       (*eDiagHistoryAbsolute*)
       1002:
         #Data.Parameter.Diag_History_Absolute.Power_Up_Counter.%B3:= #arrRecord[6];
         #Data.Parameter.Diag_History_Absolute.Power_Up_Counter.%B2:= #arrRecord[7];
         #Data.Parameter.Diag_History_Absolute.Power_Up_Counter.%B1:= #arrRecord[8];
         #Data.Parameter.Diag_History_Absolute.Power_Up_Counter.%B0:= #arrRecord[9];
         #Data.Parameter.Diag_History_Absolute.Operating_Time.%B3:= #arrRecord[10];
         #Data.Parameter.Diag_History_Absolute.Operating_Time.%B2:= #arrRecord[11];
         #Data.Parameter.Diag_History_Absolute.Operating_Time.%B1:= #arrRecord[12];
         #Data.Parameter.Diag_History_Absolute.Operating_Time.%B0:= #arrRecord[13];
         #Data.Parameter.Diag_History_Absolute.Maximum_Speed.%B3:= #arrRecord[14];
         #Data.Parameter.Diag_History_Absolute.Maximum_Speed.%B2:= #arrRecord[15];
         #Data.Parameter.Diag_History_Absolute.Maximum_Speed.%B1:= #arrRecord[16];
         #Data.Parameter.Diag_History_Absolute.Maximum_Speed.%B0:= #arrRecord[17];
         #Data.Parameter.Diag_History_Absolute.Counter_Rotation_fw.%B3:= #arrRecord[18];
         #Data.Parameter.Diag_History_Absolute.Counter_Rotation_fw.%B2:= #arrRecord[19];
         #Data.Parameter.Diag_History_Absolute.Counter_Rotation_fw.%B1:= #arrRecord[20];
         #Data.Parameter.Diag_History_Absolute.Counter_Rotation_fw.%B0:= #arrRecord[21];
         #Data.Parameter.Diag_History_Absolute.Counter_Rotation_bw.%B3:= #arrRecord[22];
         #Data.Parameter.Diag_History_Absolute.Counter_Rotation_bw.%B2:= #arrRecord[23];
         #Data.Parameter.Diag_History_Absolute.Counter_Rotation_bw.%B1:= #arrRecord[24];
         #Data.Parameter.Diag_History_Absolute.Counter_Rotation_bw.%B0:= #arrRecord[25];
         #Data.Parameter.Diag_History_Absolute.Counter_Rotation_alt.%B3:= #arrRecord[26];
         #Data.Parameter.Diag_History_Absolute.Counter_Rotation_alt.%B2:= #arrRecord[27];
         #Data.Parameter.Diag_History_Absolute.Counter_Rotation_alt.%B1:= #arrRecord[28];
         #Data.Parameter.Diag_History_Absolute.Counter_Rotation_alt.%B0:= #arrRecord[29];
         #Data.Parameter.Diag_History_Absolute.Counter_Motion.%B3:= #arrRecord[30];
         #Data.Parameter.Diag_History_Absolute.Counter_Motion.%B2:= #arrRecord[31];
         #Data.Parameter.Diag_History_Absolute.Counter_Motion.%B1:= #arrRecord[32];
         #Data.Parameter.Diag_History_Absolute.Counter_Motion.%B0:= #arrRecord[33];
         #Data.Parameter.Diag_History_Absolute.Reserved.%B3:= #arrRecord[34];
         #Data.Parameter.Diag_History_Absolute.Reserved.%B2:= #arrRecord[35];
         #Data.Parameter.Diag_History_Absolute.Reserved.%B1:= #arrRecord[36];
         #Data.Parameter.Diag_History_Absolute.Reserved.%B0:= #arrRecord[37];
         #Data.Parameter.Diag_History_Absolute.LED_Current_Maximum.%B3:= #arrRecord[38];
         #Data.Parameter.Diag_History_Absolute.LED_Current_Maximum.%B2:= #arrRecord[39];
         #Data.Parameter.Diag_History_Absolute.LED_Current_Maximum.%B1:= #arrRecord[40];
         #Data.Parameter.Diag_History_Absolute.LED_Current_Maximum.%B0:= #arrRecord[41];
         #Data.Parameter.Diag_History_Absolute.LED_Current_Minimum.%B3:= #arrRecord[42];
         #Data.Parameter.Diag_History_Absolute.LED_Current_Minimum.%B2:= #arrRecord[43];
         #Data.Parameter.Diag_History_Absolute.LED_Current_Minimum.%B1:= #arrRecord[44];
         #Data.Parameter.Diag_History_Absolute.LED_Current_Minimum.%B0:= #arrRecord[45];
         #Data.Parameter.Diag_History_Absolute.Voltage_Maximum.%B3:= #arrRecord[46];
         #Data.Parameter.Diag_History_Absolute.Voltage_Maximum.%B2:= #arrRecord[47];
         #Data.Parameter.Diag_History_Absolute.Voltage_Maximum.%B1:= #arrRecord[48];
         #Data.Parameter.Diag_History_Absolute.Voltage_Maximum.%B0:= #arrRecord[49];   
         #Data.Parameter.Diag_History_Absolute.Temperatur_Maximum.%B3:= #arrRecord[50];
         #Data.Parameter.Diag_History_Absolute.Temperatur_Maximum.%B2:= #arrRecord[51];
         #Data.Parameter.Diag_History_Absolute.Temperatur_Maximum.%B1:= #arrRecord[52];
         #Data.Parameter.Diag_History_Absolute.Temperatur_Maximum.%B0:= #arrRecord[53];
         #Data.Parameter.Diag_History_Absolute.Temperature_Minimum.%B3:= #arrRecord[54];
         #Data.Parameter.Diag_History_Absolute.Temperature_Minimum.%B2:= #arrRecord[55];
         #Data.Parameter.Diag_History_Absolute.Temperature_Minimum.%B1:= #arrRecord[56];
         #Data.Parameter.Diag_History_Absolute.Temperature_Minimum.%B0:= #arrRecord[57];

       (*eDiagHistoryRelative*)
       1003:
         #Data.Parameter.Diag_History_Relative.Power_Up_Counter.%B3:= #arrRecord[6];
         #Data.Parameter.Diag_History_Relative.Power_Up_Counter.%B2:= #arrRecord[7];
         #Data.Parameter.Diag_History_Relative.Power_Up_Counter.%B1:= #arrRecord[8];
         #Data.Parameter.Diag_History_Relative.Power_Up_Counter.%B0:= #arrRecord[9];
         #Data.Parameter.Diag_History_Relative.Operating_Time.%B3:= #arrRecord[10];
         #Data.Parameter.Diag_History_Relative.Operating_Time.%B2:= #arrRecord[11];
         #Data.Parameter.Diag_History_Relative.Operating_Time.%B1:= #arrRecord[12];
         #Data.Parameter.Diag_History_Relative.Operating_Time.%B0:= #arrRecord[13];
         #Data.Parameter.Diag_History_Relative.Maximum_Speed.%B3:= #arrRecord[14];
         #Data.Parameter.Diag_History_Relative.Maximum_Speed.%B2:= #arrRecord[15];
         #Data.Parameter.Diag_History_Relative.Maximum_Speed.%B1:= #arrRecord[16];
         #Data.Parameter.Diag_History_Relative.Maximum_Speed.%B0:= #arrRecord[17];
         #Data.Parameter.Diag_History_Relative.Counter_Rotation_fw.%B3:= #arrRecord[18];
         #Data.Parameter.Diag_History_Relative.Counter_Rotation_fw.%B2:= #arrRecord[19];
         #Data.Parameter.Diag_History_Relative.Counter_Rotation_fw.%B1:= #arrRecord[20];
         #Data.Parameter.Diag_History_Relative.Counter_Rotation_fw.%B0:= #arrRecord[21];
         #Data.Parameter.Diag_History_Relative.Counter_Rotation_bw.%B3:= #arrRecord[22];
         #Data.Parameter.Diag_History_Relative.Counter_Rotation_bw.%B2:= #arrRecord[23];
         #Data.Parameter.Diag_History_Relative.Counter_Rotation_bw.%B1:= #arrRecord[24];
         #Data.Parameter.Diag_History_Relative.Counter_Rotation_bw.%B0:= #arrRecord[25];
         #Data.Parameter.Diag_History_Relative.Counter_Rotation_alt.%B3:= #arrRecord[26];
         #Data.Parameter.Diag_History_Relative.Counter_Rotation_alt.%B2:= #arrRecord[27];
         #Data.Parameter.Diag_History_Relative.Counter_Rotation_alt.%B1:= #arrRecord[28];
         #Data.Parameter.Diag_History_Relative.Counter_Rotation_alt.%B0:= #arrRecord[29];
         #Data.Parameter.Diag_History_Relative.Counter_Motion.%B3:= #arrRecord[30];
         #Data.Parameter.Diag_History_Relative.Counter_Motion.%B2:= #arrRecord[31];
         #Data.Parameter.Diag_History_Relative.Counter_Motion.%B1:= #arrRecord[32];
         #Data.Parameter.Diag_History_Relative.Counter_Motion.%B0:= #arrRecord[33];
         #Data.Parameter.Diag_History_Relative.Reserved.%B3:= #arrRecord[34];
         #Data.Parameter.Diag_History_Relative.Reserved.%B2:= #arrRecord[35];
         #Data.Parameter.Diag_History_Relative.Reserved.%B1:= #arrRecord[36];
         #Data.Parameter.Diag_History_Relative.Reserved.%B0:= #arrRecord[37];
         #Data.Parameter.Diag_History_Relative.LED_Current_Maximum.%B3:= #arrRecord[38];
         #Data.Parameter.Diag_History_Relative.LED_Current_Maximum.%B2:= #arrRecord[39];
         #Data.Parameter.Diag_History_Relative.LED_Current_Maximum.%B1:= #arrRecord[40];
         #Data.Parameter.Diag_History_Relative.LED_Current_Maximum.%B0:= #arrRecord[41];
         #Data.Parameter.Diag_History_Relative.LED_Current_Minimum.%B3:= #arrRecord[42];
         #Data.Parameter.Diag_History_Relative.LED_Current_Minimum.%B2:= #arrRecord[43];
         #Data.Parameter.Diag_History_Relative.LED_Current_Minimum.%B1:= #arrRecord[44];
         #Data.Parameter.Diag_History_Relative.LED_Current_Minimum.%B0:= #arrRecord[45];
         #Data.Parameter.Diag_History_Relative.Voltage_Maximum.%B3:= #arrRecord[46];
         #Data.Parameter.Diag_History_Relative.Voltage_Maximum.%B2:= #arrRecord[47];
         #Data.Parameter.Diag_History_Relative.Voltage_Maximum.%B1:= #arrRecord[48];
         #Data.Parameter.Diag_History_Relative.Voltage_Maximum.%B0:= #arrRecord[49];   
         #Data.Parameter.Diag_History_Relative.Temperatur_Maximum.%B3:= #arrRecord[50];
         #Data.Parameter.Diag_History_Relative.Temperatur_Maximum.%B2:= #arrRecord[51];
         #Data.Parameter.Diag_History_Relative.Temperatur_Maximum.%B1:= #arrRecord[52];
         #Data.Parameter.Diag_History_Relative.Temperatur_Maximum.%B0:= #arrRecord[53];
         #Data.Parameter.Diag_History_Relative.Temperature_Minimum.%B3:= #arrRecord[54];
         #Data.Parameter.Diag_History_Relative.Temperature_Minimum.%B2:= #arrRecord[55];
         #Data.Parameter.Diag_History_Relative.Temperature_Minimum.%B1:= #arrRecord[56];
         #Data.Parameter.Diag_History_Relative.Temperature_Minimum.%B0:= #arrRecord[57];

       (*eDiagHistErrCounter*)
       1004:
         FOR #iIndex:= 0 TO 15 DO
           #Data.Parameter.Diag_Hist_Err_Counter[#iIndex].%B1:= #arrRecord[6 + 2 * #iIndex];
           #Data.Parameter.Diag_Hist_Err_Counter[#iIndex].%B0:= #arrRecord[7 + 2 * #iIndex];
         END_FOR;

       (*eSpeedCalculation*)
       1005:
         #Data.Parameter.Speed_Calculation.Control.%B1:= #arrRecord[6];
         #Data.Parameter.Speed_Calculation.Control.%B0:= #arrRecord[7];
         #Data.Parameter.Speed_Calculation.Velocity_Measuring_Unit.%B1:= #arrRecord[8];
         #Data.Parameter.Speed_Calculation.Velocity_Measuring_Unit.%B0:= #arrRecord[9];
         #Data.Parameter.Speed_Calculation.Update_Time_Tu.%B1:= #arrRecord[10];
         #Data.Parameter.Speed_Calculation.Update_Time_Tu.%B0:= #arrRecord[11];
         #Data.Parameter.Speed_Calculation.Update_Time_Ti.%B1:= #arrRecord[12];
         #Data.Parameter.Speed_Calculation.Update_Time_Ti.%B0:= #arrRecord[13];
         #Data.Parameter.Speed_Calculation.Upper_Limit.%B1:= #arrRecord[14];
         #Data.Parameter.Speed_Calculation.Upper_Limit.%B0:= #arrRecord[15];
         #Data.Parameter.Speed_Calculation.Lower_Limit.%B1:= #arrRecord[16];
         #Data.Parameter.Speed_Calculation.Lower_Limit.%B0:= #arrRecord[17];     

       (*eTemperatureLimits*)
       1006:
         #Data.Parameter.Temperature_Limits.Lower_Limit.%B1:= #arrRecord[6];
         #Data.Parameter.Temperature_Limits.Lower_Limit.%B0:= #arrRecord[7];
         #Data.Parameter.Temperature_Limits.Upper_Limit.%B1:= #arrRecord[8];
         #Data.Parameter.Temperature_Limits.Upper_Limit.%B0:= #arrRecord[9];   

       (*eVoltageLimits*)
       1007:
         #Data.Parameter.Voltage_Limits.Lower_Limit.%B1:= #arrRecord[6];
         #Data.Parameter.Voltage_Limits.Lower_Limit.%B0:= #arrRecord[7];
         #Data.Parameter.Voltage_Limits.Upper_Limit.%B1:= #arrRecord[8];
         #Data.Parameter.Voltage_Limits.Upper_Limit.%B0:= #arrRecord[9];   

       (*eScalingParameters*)
       1009: 
         #Data.Parameter.Scaling_Parameters.ES_Functionality.%B3:= #arrRecord[6];
         #Data.Parameter.Scaling_Parameters.ES_Functionality.%B2:= #arrRecord[7];
         #Data.Parameter.Scaling_Parameters.ES_Functionality.%B1:= #arrRecord[8];
         #Data.Parameter.Scaling_Parameters.ES_Functionality.%B0:= #arrRecord[9];
         #Data.Parameter.Scaling_Parameters.Input_CNR_N.%B3:= #arrRecord[10];
         #Data.Parameter.Scaling_Parameters.Input_CNR_N.%B2:= #arrRecord[11];
         #Data.Parameter.Scaling_Parameters.Input_CNR_N.%B1:= #arrRecord[12];
         #Data.Parameter.Scaling_Parameters.Input_CNR_N.%B0:= #arrRecord[13];
         #Data.Parameter.Scaling_Parameters.Input_CNR_D.%B3:= #arrRecord[14];
         #Data.Parameter.Scaling_Parameters.Input_CNR_D.%B2:= #arrRecord[15];
         #Data.Parameter.Scaling_Parameters.Input_CNR_D.%B1:= #arrRecord[16];
         #Data.Parameter.Scaling_Parameters.Input_CNR_D.%B0:= #arrRecord[17];
         #Data.Parameter.Scaling_Parameters.Input_CMR.%B3:= #arrRecord[18];
         #Data.Parameter.Scaling_Parameters.Input_CMR.%B2:= #arrRecord[19];
         #Data.Parameter.Scaling_Parameters.Input_CMR.%B1:= #arrRecord[20];
         #Data.Parameter.Scaling_Parameters.Input_CMR.%B0:= #arrRecord[21];
         #Data.Parameter.Scaling_Parameters.Range_Offset.%B3:= #arrRecord[22];
         #Data.Parameter.Scaling_Parameters.Range_Offset.%B2:= #arrRecord[23];
         #Data.Parameter.Scaling_Parameters.Range_Offset.%B1:= #arrRecord[24];
         #Data.Parameter.Scaling_Parameters.Range_Offset.%B0:= #arrRecord[25];
         #Data.Parameter.Scaling_Parameters.PMR_Shift.%B3:= #arrRecord[26];
         #Data.Parameter.Scaling_Parameters.PMR_Shift.%B2:= #arrRecord[27];
         #Data.Parameter.Scaling_Parameters.PMR_Shift.%B1:= #arrRecord[28];
         #Data.Parameter.Scaling_Parameters.PMR_Shift.%B0:= #arrRecord[29];
         #Data.Parameter.Scaling_Parameters.Output_CNR_N.%B3:= #arrRecord[30];
         #Data.Parameter.Scaling_Parameters.Output_CNR_N.%B2:= #arrRecord[31];
         #Data.Parameter.Scaling_Parameters.Output_CNR_N.%B1:= #arrRecord[32];
         #Data.Parameter.Scaling_Parameters.Output_CNR_N.%B0:= #arrRecord[33];
         #Data.Parameter.Scaling_Parameters.Output_CNR_D.%B3:= #arrRecord[34];
         #Data.Parameter.Scaling_Parameters.Output_CNR_D.%B2:= #arrRecord[35];
         #Data.Parameter.Scaling_Parameters.Output_CNR_D.%B1:= #arrRecord[36];
         #Data.Parameter.Scaling_Parameters.Output_CNR_D.%B0:= #arrRecord[37];
         #Data.Parameter.Scaling_Parameters.Output_CMR.%B3:= #arrRecord[38];
         #Data.Parameter.Scaling_Parameters.Output_CMR.%B2:= #arrRecord[39];
         #Data.Parameter.Scaling_Parameters.Output_CMR.%B1:= #arrRecord[40];
         #Data.Parameter.Scaling_Parameters.Output_CMR.%B0:= #arrRecord[41];
         #Data.Parameter.Scaling_Parameters.Out_CPR_Integer.%B3:= #arrRecord[42];
         #Data.Parameter.Scaling_Parameters.Out_CPR_Integer.%B2:= #arrRecord[43];
         #Data.Parameter.Scaling_Parameters.Out_CPR_Integer.%B1:= #arrRecord[44];
         #Data.Parameter.Scaling_Parameters.Out_CPR_Integer.%B0:= #arrRecord[45];
         #Data.Parameter.Scaling_Parameters.Out_CPR_Fract.%B3:= #arrRecord[46];
         #Data.Parameter.Scaling_Parameters.Out_CPR_Fract.%B2:= #arrRecord[47];
         #Data.Parameter.Scaling_Parameters.Out_CPR_Fract.%B1:= #arrRecord[48];
         #Data.Parameter.Scaling_Parameters.Out_CPR_Fract.%B0:= #arrRecord[49];

       (*eOperationTest1*)
       1010:
         #Data.Parameter.Operation_Test_1.%B1:= #arrRecord[6];
         #Data.Parameter.Operation_Test_1.%B0:= #arrRecord[7];

       (*eMACIDPort1*)
       1011:
         FOR #iIndex:= 0 TO 5 DO
           #Data.Parameter.MAC_ID_Port_1[#iIndex]:= #arrRecord[6 + #iIndex];
         END_FOR;

       (*eMACIDPort2*)
       1012:
         FOR #iIndex:= 0 TO 5 DO
           #Data.Parameter.MAC_ID_Port_2[#iIndex]:= #arrRecord[6 + #iIndex];
         END_FOR;

       (*eVersionFWFPGA*)
       1013:
         #Data.Parameter.Version_FW_FPGA.%B3:= #arrRecord[6];
         #Data.Parameter.Version_FW_FPGA.%B2:= #arrRecord[7];
         #Data.Parameter.Version_FW_FPGA.%B1:= #arrRecord[8];
         #Data.Parameter.Version_FW_FPGA.%B0:= #arrRecord[9];

       (*eTemperature*)
       1014:
         #Data.Parameter.Temperature.%B1:= #arrRecord[6];  
         #Data.Parameter.Temperature.%B0:= #arrRecord[7];  

       (*eStationName*)
       61000:
         Chars_TO_Strg(Chars:= #arrRecord, pChars:= 6, Cnt:= BYTE_TO_UINT(#arrRecord[5]), Strg=>#Data.Parameter.Station_Name);

       (*eStationIP*)
       61001:
         FOR #iIndex:= 0 TO 3 DO
           #Data.Parameter.Station_IP[#iIndex]:= #arrRecord[6 + #iIndex];
         END_FOR;

       (*eStationMACID*)
       61002:
         FOR #iIndex:= 0 TO 5 DO
           #Data.Parameter.Station_MAC_ID[#iIndex]:= #arrRecord[6 + #iIndex];
         END_FOR;

       (*eStationGateway*)
       61003:
         FOR #iIndex:= 0 TO 3 DO
           #Data.Parameter.Station_Gateway[#iIndex]:= #arrRecord[6 + #iIndex];
         END_FOR;

       (*eStationSubnet*)
       61004:
         FOR #iIndex:= 0 TO 3 DO
           #Data.Parameter.Station_Subnet[#iIndex]:= #arrRecord[6 + #iIndex];
         END_FOR;

       (*ePresetValue*)
       65000:
         #Data.Parameter.Preset_Value.%B3:= #arrRecord[6];
         #Data.Parameter.Preset_Value.%B2:= #arrRecord[7];
         #Data.Parameter.Preset_Value.%B1:= #arrRecord[8];
         #Data.Parameter.Preset_Value.%B0:= #arrRecord[9];

       (*eOperatingStatus*)
       65001:
         #Data.Parameter.Operating_Status.Header.%B3:= #arrRecord[6];
         #Data.Parameter.Operating_Status.Header.%B2:= #arrRecord[7];
         #Data.Parameter.Operating_Status.Header.%B1:= #arrRecord[8];
         #Data.Parameter.Operating_Status.Header.%B0:= #arrRecord[9];
         #Data.Parameter.Operating_Status.Operating_Status.%B3:= #arrRecord[10];
         #Data.Parameter.Operating_Status.Operating_Status.%B2:= #arrRecord[11];
         #Data.Parameter.Operating_Status.Operating_Status.%B1:= #arrRecord[12];
         #Data.Parameter.Operating_Status.Operating_Status.%B0:= #arrRecord[13];
         #Data.Parameter.Operating_Status.Faults.%B3:= #arrRecord[14];
         #Data.Parameter.Operating_Status.Faults.%B2:= #arrRecord[15];
         #Data.Parameter.Operating_Status.Faults.%B1:= #arrRecord[16];
         #Data.Parameter.Operating_Status.Faults.%B0:= #arrRecord[17];
         #Data.Parameter.Operating_Status.Supported_Faults.%B3:= #arrRecord[18];
         #Data.Parameter.Operating_Status.Supported_Faults.%B2:= #arrRecord[19];
         #Data.Parameter.Operating_Status.Supported_Faults.%B1:= #arrRecord[20];
         #Data.Parameter.Operating_Status.Supported_Faults.%B0:= #arrRecord[21];
         #Data.Parameter.Operating_Status.Warnings.%B3:= #arrRecord[22];
         #Data.Parameter.Operating_Status.Warnings.%B2:= #arrRecord[23];
         #Data.Parameter.Operating_Status.Warnings.%B1:= #arrRecord[24];
         #Data.Parameter.Operating_Status.Warnings.%B0:= #arrRecord[25];
         #Data.Parameter.Operating_Status.Supported_Warnings.%B3:= #arrRecord[26];
         #Data.Parameter.Operating_Status.Supported_Warnings.%B2:= #arrRecord[27];
         #Data.Parameter.Operating_Status.Supported_Warnings.%B1:= #arrRecord[28];
         #Data.Parameter.Operating_Status.Supported_Warnings.%B0:= #arrRecord[29];
         #Data.Parameter.Operating_Status.Encoder_Profile_Version.%B3:= #arrRecord[30];
         #Data.Parameter.Operating_Status.Encoder_Profile_Version.%B2:= #arrRecord[31];
         #Data.Parameter.Operating_Status.Encoder_Profile_Version.%B1:= #arrRecord[32];
         #Data.Parameter.Operating_Status.Encoder_Profile_Version.%B0:= #arrRecord[33];
         #Data.Parameter.Operating_Status.Operating_Time.%B3:= #arrRecord[34];
         #Data.Parameter.Operating_Status.Operating_Time.%B2:= #arrRecord[35];
         #Data.Parameter.Operating_Status.Operating_Time.%B1:= #arrRecord[36];
         #Data.Parameter.Operating_Status.Operating_Time.%B0:= #arrRecord[37];
         #Data.Parameter.Operating_Status.Offset_Value.%B3:= #arrRecord[38];
         #Data.Parameter.Operating_Status.Offset_Value.%B2:= #arrRecord[39];
         #Data.Parameter.Operating_Status.Offset_Value.%B1:= #arrRecord[40];
         #Data.Parameter.Operating_Status.Offset_Value.%B0:= #arrRecord[41];
         #Data.Parameter.Operating_Status.CPR.%B3:= #arrRecord[42];
         #Data.Parameter.Operating_Status.CPR.%B2:= #arrRecord[43];
         #Data.Parameter.Operating_Status.CPR.%B1:= #arrRecord[44];
         #Data.Parameter.Operating_Status.CPR.%B0:= #arrRecord[45];
         #Data.Parameter.Operating_Status.CMR.%B3:= #arrRecord[46];
         #Data.Parameter.Operating_Status.CMR.%B2:= #arrRecord[47];
         #Data.Parameter.Operating_Status.CMR.%B1:= #arrRecord[48];
         #Data.Parameter.Operating_Status.CMR.%B0:= #arrRecord[49];
         #Data.Parameter.Operating_Status.Velocity_Measuring_Unit.%B3:= #arrRecord[50];
         #Data.Parameter.Operating_Status.Velocity_Measuring_Unit.%B2:= #arrRecord[51];
         #Data.Parameter.Operating_Status.Velocity_Measuring_Unit.%B1:= #arrRecord[52];
         #Data.Parameter.Operating_Status.Velocity_Measuring_Unit.%B0:= #arrRecord[53];
     ELSE
       #stTempErrorCode.nBlockError:= 16#0002; (*Error: Internal error*)
     END_CASE;
     #iStep:= 9; (*Action permormed / Next command*)
   END_IF;


   (*======================== ACTION PERFORMED / NEXT COMMAND (STEP 9) =========================*)
   IF #iStep = 9 THEN
     #iCommandIndex:= #iCommandIndex + 1;

     (*Job done*)
     IF (#iCommandIndex > 31) OR (#arrCommandQueue[#iCommandIndex].iPNU <= 0) THEN
       #Done:= true;
       #Busy:= false;
       #bBusyMem:= false;
       #Error:= false;
       #iStep:= 0;

     (*Next command*)
     ELSE
       #iStep:= 4; (*Check communication status*)
     END_IF;
   END_IF;
END_FUNCTION_BLOCK

FUNCTION "Conveyors_Transfer" : Void   // FC24, SCL
{ S7_Optimized_Access := 'TRUE' }
VERSION : 0.1
// stored: AutoNumber true, IsIECCheckEnabled false, SetENOAutomatically false, UDAEnableTagReadback false
   VAR_TEMP
      i : Int;
   END_VAR
BEGIN
   //ID OF THE VTD CONVEYOR
   IF "Control_DB".VTD_Control.Current_Level = 0 THEN
       "Settings_DB".ECnv_Settings.ID := 120001;
       "Settings_DB".ECnv_Settings.Cnv_Level := 0;
   ELSIF "Control_DB".VTD_Control.Current_Level = 1 THEN
       "Settings_DB".ECnv_Settings.ID := 120101;
       "Settings_DB".ECnv_Settings.Cnv_Level := 1;
   ELSIF "Control_DB".VTD_Control.Current_Level = 2 THEN
       "Settings_DB".ECnv_Settings.ID := 120201;
       "Settings_DB".ECnv_Settings.Cnv_Level := 2;
   ELSIF "Control_DB".VTD_Control.Current_Level = 3 THEN
       "Settings_DB".ECnv_Settings.ID := 120301;
       "Settings_DB".ECnv_Settings.Cnv_Level := 3;
   ELSE
       "Settings_DB".ECnv_Settings.ID := 129901;
       "Settings_DB".ECnv_Settings.Cnv_Level := 99;
   END_IF;

   REGION READY TO RECEIVE
       //EXTRACTOR CONVEYOR
       "Control_DB".ECnv_Control.Instruction.Inbound_Ready :=
       ("Settings_DB".ECnv_Settings.ID = 120001 OR
       "Settings_DB".ECnv_Settings.ID = 120101 OR
       "Settings_DB".ECnv_Settings.ID = 120201 OR
       "Settings_DB".ECnv_Settings.ID = 120301)
       AND NOT "Control_DB".ECnv_Control.Cnv_Occupied AND NOT "Control_DB".ECnv_Control.Instruction.Outbound_Ready AND
       ("Control_DB".ECnv_Control.Mode = 2 OR "Control_DB".ECnv_Control.Mode = 3);

       //BUFFER CONVEYORS
       FOR #i := 1 TO 3 DO
           "Control_DB".LCnv_Control[#i].Instruction.Inbound_Ready :=
           NOT "Control_DB".LCnv_Control[#i].Running AND
           NOT "Control_DB".LCnv_Control[#i].Cnv_Occupied AND NOT "Control_DB".LCnv_Control[#i].Instruction.Outbound_Ready AND
           ("Control_DB".LCnv_Control[#i].Mode = 2 OR "Control_DB".LCnv_Control[#i].Mode = 3);
       END_FOR;

       //POPUP CONVEYORS
       FOR #i := 1 TO 4 DO
           "Control_DB".PopUp_Cnv[#i].Instruction.Inbound_Ready :=
           NOT "Control_DB".PopUp_Cnv[#i].Running AND
           NOT "Control_DB".PopUp_Cnv[#i].Cnv_Occupied AND NOT "Control_DB".PopUp_Cnv[#i].Instruction.Outbound_Ready AND
           ("Control_DB".PopUp_Cnv[#i].Mode = 2 OR "Control_DB".PopUp_Cnv[#i].Mode = 3);
       END_FOR;

       //INBOUND CONVEYOR
       "Control_DB".Inbound_Cnv.Instruction.Inbound_Ready := NOT "Control_DB".Inbound_Cnv.Cnv_Occupied;

       //OUTBOUND CONVEYOR
       "Control_DB".Outbound_Cnv.Instruction.Inbound_Ready :=
       NOT "Control_DB".Outbound_Cnv.Running AND
       NOT "Control_DB".Outbound_Cnv.Cnv_Occupied AND NOT "Control_DB".Outbound_Cnv.Instruction.Outbound_Ready AND
       ("Control_DB".Outbound_Cnv.Mode = 2 OR "Control_DB".Outbound_Cnv.Mode = 3);

       //PICK CONVEYOR
       "Control_DB".Pick_Station.Instruction.Inbound_Ready :=
       NOT "Control_DB".Pick_Station.Running AND
       NOT "Control_DB".Pick_Station.Cnv_Occupied AND NOT "Control_DB".Pick_Station.Instruction.Outbound_Ready AND
       ("Control_DB".Pick_Station.Mode = 2 OR "Control_DB".Pick_Station.Mode = 3);
   END_REGION

   REGION READY TO SEND
       //EXTRACTOR CONVEYOR
       "Control_DB".ECnv_Control.Instruction.Outbound_Ready :=
       (("Settings_DB".ECnv_Settings.ID = 120001 AND "Control_DB".ECnv_Control.Cnv_Occupied AND
       NOT "Control_DB".PopUp_Cnv[2].Cnv_Occupied AND ("Control_DB".PopUp_Cnv[2].Mode = 2 OR "Control_DB".PopUp_Cnv[2].Mode = 3)
       AND NOT "Control_DB".PopUp_Cnv[2].Error)
       OR
       ("Settings_DB".ECnv_Settings.ID = 120101 AND "Control_DB".ECnv_Control.Cnv_Occupied AND
       NOT "Control_DB".LCnv_Control[1].Cnv_Occupied AND ("Control_DB".LCnv_Control[1].Mode = 2 OR "Control_DB".LCnv_Control[1].Mode = 3)
       AND NOT "Control_DB".LCnv_Control[1].Error)
       OR
       ("Settings_DB".ECnv_Settings.ID = 120201 AND "Control_DB".ECnv_Control.Cnv_Occupied AND
       NOT "Control_DB".LCnv_Control[2].Cnv_Occupied AND ("Control_DB".LCnv_Control[2].Mode = 2 OR "Control_DB".LCnv_Control[2].Mode = 3)
       AND NOT "Control_DB".LCnv_Control[2].Error)
       OR
       ("Settings_DB".ECnv_Settings.ID = 120301 AND "Control_DB".ECnv_Control.Cnv_Occupied AND
       NOT "Control_DB".LCnv_Control[3].Cnv_Occupied AND ("Control_DB".LCnv_Control[3].Mode = 2 OR "Control_DB".LCnv_Control[3].Mode = 3)
       AND NOT "Control_DB".LCnv_Control[3].Error));

       //BUFFER CONVEYORS
       FOR #i := 1 TO 3 DO
           "Control_DB".LCnv_Control[#i].Instruction.Outbound_Ready :=
           "Control_DB".ECnv_Control.Instruction.Inbound_Ready AND
           "Control_DB".VTD_Control.Current_Level = #i AND
           NOT "Control_DB".LCnv_Control[#i].Instruction.Transfer_in_Progress AND
           "Control_DB".LCnv_Control[#i].Cnv_Occupied AND
           ("Control_DB".LCnv_Control[#i].Mode = 2 OR "Control_DB".LCnv_Control[#i].Mode = 3);
       END_FOR;

       //INBOUND CONVEYOR
       "Control_DB".Inbound_Cnv.Instruction.Outbound_Ready := "Control_DB".Inbound_Cnv.Cnv_Occupied;

       //POPUP CONVEYORS
       FOR #i := 1 TO 4 DO
           "Control_DB".PopUp_Cnv[#i].Instruction.Outbound_Ready :=
           ((#i = 1 AND "Control_DB".PopUp_Cnv[2].Instruction.Inbound_Ready AND "Control_DB".PopUp_Cnv[1].Inputs."Lift Up") OR
           (#i = 2 AND "Control_DB".PopUp_Cnv[2].Inputs."Lift Down" AND ("Control_DB".PopUp_Cnv[3].Instruction.Inbound_Ready OR "Control_DB".ECnv_Control.Instruction.Inbound_Ready)) OR
           (#i = 3 AND "Control_DB".PopUp_Cnv[4].Instruction.Inbound_Ready AND "Control_DB".PopUp_Cnv[3].Inputs."Lift Up") OR
           (#i = 4 AND ("Control_DB".Outbound_Cnv.Instruction.Inbound_Ready OR "Control_DB".PopUp_Cnv[1].Instruction.Inbound_Ready) AND ("Control_DB".PopUp_Cnv[4].Inputs."Lift Up" OR "Control_DB".PopUp_Cnv[4].Inputs."Lift Down"))) AND
           (*("Control_DB".VTD_Control.Current_Level = 0 AND #i = 2) AND*)
           NOT "Control_DB".PopUp_Cnv[#i].Instruction.Transfer_in_Progress AND
           "Control_DB".PopUp_Cnv[#i].Cnv_Occupied = TRUE AND
           ("Control_DB".PopUp_Cnv[#i].Mode = 2 OR "Control_DB".PopUp_Cnv[#i].Mode = 3);
       END_FOR;

       //PICK CONVEYOR
       "Control_DB".Pick_Station.Instruction.Outbound_Ready := "Control_DB".Pick_Station.Cnv_Occupied;
   END_REGION

   REGION TRANSFER IN PROGRESS FOR VTD
       "Cnv_TIP_For_VTD" :=
       ("Settings_DB".ECnv_Settings.ID = 120001 AND
       "Control_DB".PopUp_Cnv[2].Instruction.Transfer_in_Progress)
       OR
       ("Settings_DB".ECnv_Settings.ID = 120101 AND
       "Control_DB".LCnv_Control[1].Instruction.Transfer_in_Progress)
       OR
       ("Settings_DB".ECnv_Settings.ID = 120201 AND
       "Control_DB".LCnv_Control[2].Instruction.Transfer_in_Progress)
       OR
       ("Settings_DB".ECnv_Settings.ID = 120301 AND
       "Control_DB".LCnv_Control[3].Instruction.Transfer_in_Progress);
   END_REGION
END_FUNCTION

FUNCTION_BLOCK "Light_Bars"   // FB6, SCL
{ S7_Optimized_Access := 'TRUE' }
VERSION : 0.1
// stored: AutoNumber true, IsIECCheckEnabled false, IsRetainMemResEnabled false, MemoryReserve 100, SetENOAutomatically false, UDAEnableTagReadback false
   VAR_INPUT
      VTD_Mode : UInt;
      VTD_Speed : Int;
      Fault : Bool;
   END_VAR
   VAR_OUTPUT
      Animation_B1 : Byte;
      Color_B1 : Byte;
      Animation_B2 : Byte;
      Color_B2 : Byte;
      Speed_B1 : Byte;
      Speed_B2 : Byte;
   END_VAR
BEGIN
   //Commands for Light Bar

   IF #VTD_Mode = 0 AND NOT #Fault THEN // (0)Disabled = No light  
       #Animation_B1:= #Animation_B2:= 0;

   ELSIF #VTD_Mode = 1 AND #VTD_Speed = 0 AND  NOT #Fault AND NOT "SinaSpeed_VTD".EnableAxis THEN // (1)Manual= Yellow Stop
       #Animation_B1 := #Animation_B2 := 1;
       #Color_B1 := #Color_B2 := 4;

   ELSIF #VTD_Mode = 1 AND #VTD_Speed > 0 AND #VTD_Speed <= 33 AND  NOT #Fault AND "SinaSpeed_VTD".EnableAxis THEN // (1)Manual= Yellow until 33%
       #Animation_B1 := #Animation_B2 := 2;
       #Speed_B1 := #Speed_B2 := 2;
       #Color_B1 := #Color_B2 := 4;

   ELSIF #VTD_Mode = 1 AND #VTD_Speed > 33 AND #VTD_Speed <= 100 AND  NOT #Fault THEN // (1)Manual= Yellow until 66%
       #Animation_B1 := #Animation_B2 := 2;
       #Speed_B1 := #Speed_B2 := 0;
       #Color_B1 := #Color_B2 := 4;

   // ELSIF #VTD_Mode = 1 AND #VTD_Speed > 66 AND #VTD_Speed <= 100 AND  NOT #Fault THEN // (1)Manual= Yellow until 100%
   //     #Animation_B1 := #Animation_B2 := 2;
   //     #Speed_B1 := #Speed_B2 := 1;
   //     #Color_B1 := #Color_B2 := 4;

   ELSIF #VTD_Mode = 2 AND #VTD_Speed = 0 AND  NOT #Fault AND NOT "SinaSpeed_VTD".EnableAxis THEN // (2)Semi-auto = Blue Stop
       #Animation_B1 := #Animation_B2 := 1;
       #Color_B1 := #Color_B2 := 9;
       #Speed_B1 := #Speed_B2 := 0;

   ELSIF #VTD_Mode = 2 AND #VTD_Speed > 0 AND #VTD_Speed <= 33 AND  NOT #Fault AND "SinaSpeed_VTD".EnableAxis THEN // (2)Semi-auto = Blue until 33%
       #Animation_B1 := #Animation_B2 := 2;
       #Speed_B1 := #Speed_B2 := 2;
       #Color_B1 := #Color_B2 := 9;

   ELSIF #VTD_Mode = 2 AND #VTD_Speed > 33 AND #VTD_Speed <= 100 AND  NOT #Fault THEN // (2)Semi-auto = Blue until 66%
       #Animation_B1 := #Animation_B2 := 2;
       #Speed_B1 := #Speed_B2 := 0;
       #Color_B1 := #Color_B2 := 9;

   // ELSIF #VTD_Mode = 2 AND #VTD_Speed > 66 AND #VTD_Speed <= 100 AND  NOT #Fault THEN // (2)Semi-auto = Blue until 100%
   //     #Animation_B1 := #Animation_B2 := 2;
   //     #Speed_B1 := #Speed_B2 := 1;
   //     #Color_B1 := #Color_B2 := 9;

   ELSIF #VTD_Mode = 3 AND #VTD_Speed = 0 AND  NOT #Fault AND NOT "SinaSpeed_VTD".EnableAxis THEN // (3)Auto = Green Stop
       #Animation_B1 := #Animation_B2 := 1;
       #Color_B1 := #Color_B2 := 0;

   ELSIF #VTD_Mode = 3 AND #VTD_Speed > 0 AND #VTD_Speed <= 33 AND  NOT #Fault AND "SinaSpeed_VTD".EnableAxis THEN // (3)Auto = Green until 33%
       #Animation_B1 := #Animation_B2 := 2;
       #Speed_B1 := #Speed_B2 := 2;
       #Color_B1 := #Color_B2 := 0;

   ELSIF #VTD_Mode = 3 AND #VTD_Speed > 33 AND #VTD_Speed <= 100 AND  NOT #Fault THEN // (3)Auto = Green until 66%
       #Animation_B1 := #Animation_B2 := 2;
       #Speed_B1 := #Speed_B2 := 0;
       #Color_B1 := #Color_B2 := 0;

   // ELSIF #VTD_Mode = 3 AND #VTD_Speed > 66 AND #VTD_Speed <= 100 AND  NOT #Fault THEN // (3)Auto = Green until 100%
   //     #Animation_B1 := #Animation_B2 := 2;
   //     #Speed_B1 := #Speed_B2 := 1;
   //     #Color_B1 := #Color_B2 := 0;

   ELSIF #VTD_Mode = 4 AND #VTD_Speed = 0 AND  NOT #Fault THEN // (4)Tech = Orange Stop
       #Animation_B1 := #Animation_B2 := 1;
       #Color_B1 := #Color_B2 := 2;

   ELSIF #VTD_Mode = 4 AND #VTD_Speed > 0 AND #VTD_Speed <= 33 AND  NOT #Fault THEN // (4)Tech = Orange until 33%
       #Animation_B1 := #Animation_B2 := 2;
       #Speed_B1 := #Speed_B2 := 2;
       #Color_B1 := #Color_B2 := 2;

   ELSIF #VTD_Mode = 4 AND #VTD_Speed > 33 AND #VTD_Speed <= 66 AND  NOT #Fault THEN // (4)Tech = Orange until 66%
       #Animation_B1 := #Animation_B2 := 2;
       #Speed_B1 := #Speed_B2 := 0;
       #Color_B1 := #Color_B2 := 2;

   ELSIF #VTD_Mode = 4 AND #VTD_Speed > 66 AND #VTD_Speed <= 100 AND  NOT #Fault THEN // (4)Tech = Orange until 100%
       #Animation_B1 := #Animation_B2 := 2;
       #Speed_B1 := #Speed_B2 := 1;
       #Color_B1 := #Color_B2 := 2;

   ELSIF #VTD_Mode = 5 AND #VTD_Speed = 0 AND  NOT #Fault THEN // (5)Maintenance = White Stop
       #Animation_B1 := #Animation_B2 := 1;
       #Color_B1 := #Color_B2 := 19;

   ELSIF #VTD_Mode = 5 AND #VTD_Speed > 0 AND #VTD_Speed <= 33 AND  NOT #Fault THEN // (5)Maintenance = White until 33%
       #Animation_B1 := #Animation_B2 := 2;
       #Speed_B1 := #Speed_B2 := 2;
       #Color_B1 := #Color_B2 := 19;

   ELSIF #VTD_Mode = 5 AND #VTD_Speed > 33 AND #VTD_Speed <= 66 AND  NOT #Fault THEN // (5)Maintenance = White until 66%
       #Animation_B1 := #Animation_B2 := 2;
       #Speed_B1 := #Speed_B2 := 0;
       #Color_B1 := #Color_B2 := 19;

   ELSIF #VTD_Mode = 5 AND #VTD_Speed > 66 AND #VTD_Speed <= 100 AND  NOT #Fault THEN // (5)Maintenance = White until 100%
       #Animation_B1 := #Animation_B2 := 2;
       #Speed_B1 := #Speed_B2 := 1;
       #Color_B1 := #Color_B2 := 19;

   ELSIF #Fault THEN // Fault = Flash Red
       #Animation_B1:= #Animation_B2 := 2;
       #Color_B1:=#Color_B2 := 1;
   END_IF;
END_FUNCTION_BLOCK

FUNCTION_BLOCK "SICK_Lector_CLV6xx_PNDP"   // FB72, SCL
TITLE = SICK Lector6xx / CLV6xx function block
{ S7_Optimized_Access := 'TRUE' }
AUTHOR : SICKAG
FAMILY : Ident
VERSION : 1.2
// This function block is used for a communication between a SICK Lector6xx / SICK CLV6xx code reader and a Siemens S7-1200/S7-1500 PLC via  PROFINET/PROFIBUS
// stored: AutoNumber false, IsIECCheckEnabled false, IsRetainMemResEnabled false, MemoryReserve 100, SetENOAutomatically false, UDAEnableTagReadback false
   VAR_INPUT
      HWInputIdent : HW_IO;   // Hardware identification number of the input module
      HWInputLength : USInt;   // Size of the input module
      HWOutputIdent : HW_IO;   // Hardware identification number of the output module
      HWOutputLength : USInt;   // Size of the output module
      CANId : USInt;   // CAN ID (0= Master / No CAN network)
      TOut : Time := T#10s;   // Time out
      Req : Bool;   // A positive edge starts the request
      TriggerOn : Bool;   // Select: Trigger On to open the reading gate via a SW-Trigger command
      TriggerOff : Bool;   // Select: Trigger Off to close the reading gate via a SW-Trigger command
      Matchcode : Bool;   // Select: Matchcode (details at #Data)
      SavePermanent : Bool;   // Select: Save permanent
      ComTest : Bool;   // Select: Communication test
      FreeCommand : Bool;   // Select: Free command (details at #Data)
   END_VAR
   VAR_OUTPUT
      RdDone : Bool;   // Positive edge: A reading result sent by the device was received
      ReqDone : Bool;   // Request done
      ReqBusy : Bool;   // Request in process
      Error : Bool;   // Error detected
      Errorcode : DWord;   // Error code (see documentation)
   END_VAR
   VAR_IN_OUT
      Data : "ST_SICK_Lector_CLV6xx";   // Command arguments and result outputs of the FB actions
   END_VAR
   VAR
      bTriggerReq { ExternalAccessible := 'False'; ExternalVisible := 'False'; ExternalWritable := 'False'} : Bool;   // Rising edge detection
      bTriggerReqMem { ExternalAccessible := 'False'; ExternalVisible := 'False'; ExternalWritable := 'False'} : Bool;   // Rising edge detection
      bTriggerDone { ExternalAccessible := 'False'; ExternalVisible := 'False'; ExternalWritable := 'False'} : Bool;   // Rising edge detection
      bTriggerDoneMem { ExternalAccessible := 'False'; ExternalVisible := 'False'; ExternalWritable := 'False'} : Bool;   // Rising edge detection
      bTriggerError { ExternalAccessible := 'False'; ExternalVisible := 'False'; ExternalWritable := 'False'} : Bool;   // Rising edge detection
      bTriggerErrorMem { ExternalAccessible := 'False'; ExternalVisible := 'False'; ExternalWritable := 'False'} : Bool;   // Rising edge detection
      bCanActive { ExternalAccessible := 'False'; ExternalVisible := 'False'; ExternalWritable := 'False'} : Bool;   // CAN-Bus active flag
      bDeviceState { ExternalAccessible := 'False'; ExternalVisible := 'False'; ExternalWritable := 'False'} : Bool;   // Current device state (True= Edit-Mode | False= Run-Mode)
      bEnforceLogout { ExternalAccessible := 'False'; ExternalVisible := 'False'; ExternalWritable := 'False'} : Bool;   // Logout enforced
      bReqBusyMem : Bool;   // Backup variable
      iStep { ExternalAccessible := 'False'; ExternalVisible := 'False'; ExternalWritable := 'False'} : USInt;   // Currrent FB step
      iCommandIndex { ExternalAccessible := 'False'; ExternalVisible := 'False'; ExternalWritable := 'False'} : Int;   // Command index
      iCommandLength { ExternalAccessible := 'False'; ExternalVisible := 'False'; ExternalWritable := 'False'} : UInt;   // Length of the command that should be send
      iRecordSize { ExternalAccessible := 'False'; ExternalVisible := 'False'; ExternalWritable := 'False'} : UInt;   // Length of the record array
      iCommandSize { ExternalAccessible := 'False'; ExternalVisible := 'False'; ExternalWritable := 'False'} : UInt;   // Length of the command array
      iReadingResultSize { ExternalAccessible := 'False'; ExternalVisible := 'False'; ExternalWritable := 'False'} : UInt;   // Length of the reading result array
      iIndex { ExternalAccessible := 'False'; ExternalVisible := 'False'; ExternalWritable := 'False'} : UInt;   // Index variable
      nTempErrorCode { ExternalAccessible := 'False'; ExternalVisible := 'False'; ExternalWritable := 'False'} : DWord;   // Temporarily error code
      nLogoutErrorCode { ExternalAccessible := 'False'; ExternalVisible := 'False'; ExternalWritable := 'False'} : DWord;   // Temporarily error code
      arrSelection { ExternalAccessible := 'False'; ExternalVisible := 'False'; ExternalWritable := 'False'} : Array[0..5] of Bool;   // input bit selection
      arrCommand { ExternalAccessible := 'False'; ExternalVisible := 'False'; ExternalWritable := 'False'} : Array[0..499] of Byte;   // Contains the transmitted CoLa command
      arrRecord { ExternalAccessible := 'False'; ExternalVisible := 'False'; ExternalWritable := 'False'} : Array[0..499] of Byte;   // Contains the received telegram
      fbTimeout { ExternalAccessible := 'False'; ExternalVisible := 'False'; ExternalWritable := 'False'; S7_SetPoint := 'True'} : TON_TIME;   // Instance: Timer on delay (Time out)
      fbCCom { ExternalAccessible := 'False'; ExternalVisible := 'False'; ExternalWritable := 'False'; S7_SetPoint := 'True'} : "SICK_CCOMM_PNDP";   // Instance: CoLa communication block
   END_VAR
   VAR_TEMP
      iTemp1 : Int;   // Temporarily variable
      iTemp2 : UDInt;   // Temporarily variable
      iTemp3 : UDInt;   // Temporarily variable
      nFncValue : DWord;   // Get/Set function value
      nFncErrorCode : Word;   // Get/Set function error code
   END_VAR
BEGIN
   (*===========================================================================================
   Name:   SICK_Lector_CLV6xx_PNDP 
   Author: SICK AG
   =============================================================================================
   Description: 
   This function block is used for a communication between a SICK Lector6xx / SICK CLV6xx
   code reader and a Siemens S7-1200/S7-1500 PLC via PROFINET/PROFIBUS.                         

   =============================================================================================
   Features:        
   - Receive reading results of the device, triggered by a command, fieldbus or by a hardware 
     switch. The content of the result can be modified in the "Output Format" option in the
     SOPAS engineeringtool.                                           
   - Open and close a reading gate (software trigger via command)
   - Set a new Matchcode evaluation condition 
   - Save all device parameters permanent                                                  
   - Communication test
   - Send a free defined CoLa-A telegram and receive the result
   - All commands can also be used in a SICK CAN-Bus network

   =============================================================================================
   Version history:
   Date       | Version | Author  | Remark
   ---------------------------------------------------------------------------------------------
   21/02/2014 | V1.0    | SICK AG | Initial version
   07/08/2014 | V1.1    | SICK AG | Replace R_TRIG function 
   24/10/2017 | V1.2    | SICK AG | Avoid initialization warnings which occurs using TIA V13 or higher
   ============================================================================================*)

   (*===================================== INITIALISATION =====================================*)
   #iRecordSize:= 500;         (*Length of the arrRecord array*)
   #iCommandSize:= 500;        (*Length of the arrCommand array*)
   #iReadingResultSize:= 200;  (*Length of the reading result array*)

   (*Rising edge detection*)
   #bTriggerReq:= #Req AND NOT #bTriggerReqMem;
   #bTriggerReqMem:= #Req;
   #bTriggerDone:= #fbCCom.ReqDone AND NOT #bTriggerDoneMem;
   #bTriggerDoneMem:= #fbCCom.ReqDone;
   #bTriggerError:= #fbCCom.Error AND NOT #bTriggerErrorMem;
   #bTriggerErrorMem:= #fbCCom.Error;

   (*Reset the read done flag every cycle*)
   #RdDone:= false;


   (*===================================== ERROR HANDLING =====================================*)
   (* bDeviceState  |  bEnforceLogout  |  Action
          FALSE     |      FALSE       |  Errorcode = Errorcode from last plc cycle
          FALSE     |      TRUE        |  Errorcode = Logout error
          TRUE      |      FALSE       |  Enforce "Logout" command
          TRUE      |      TRUE        |  Errorcode = Logout not possible + Reason*)
   IF #nTempErrorCode <>16#0000_0000 THEN

     (*Enfore "Logout" command*)
     IF #bDeviceState AND NOT #bEnforceLogout THEN
       #bEnforceLogout:= true;
       #iCommandIndex:= 11;                  (*Logout*)
       #nLogoutErrorCode:= #nTempErrorCode;  (*Save current error code*)
       #nTempErrorCode:= 16#0000_0000;       (*Clear currenr error variable*)
       #iStep:= 4;                           (*Create command*)

     (*Logout can not be ensured*)
     ELSIF #bDeviceState AND #bEnforceLogout THEN
       #Errorcode.%W1:= #nTempErrorCode.%W0;  
       #Errorcode.%W0:= 16#0017;  (*Error: Logout can not be ensured (please check the device state)*)

     (*Errorcode = Errorcode from the last plc cycle or logout error*)
     ELSE
       #Errorcode:= #nTempErrorCode;
     END_IF;

     (*Update FB status*)
     IF #nTempErrorCode <> 16#0000_0000 THEN
       #ReqDone:= false;
       #ReqBusy:= false;
       #bReqBusyMem:= false;
       #Error:= true;
       #nTempErrorCode:= 16#0000_0000;
       #nLogoutErrorCode:= 16#0000_0000;
       #iStep:= 0;
       RETURN;
     END_IF;
   END_IF;

   (*Time out detection*)
   #fbTimeout(IN:= #bReqBusyMem, PT:= #TOut);
   IF #fbTimeout.Q THEN
     #nTempErrorCode:= 16#0000_0010; (*Error: Time out*)
   END_IF;

   (*Check if a device error is detected: 'sFA XX'*)
   IF #bTriggerDone AND ((NOT #bCanActive AND
     #arrRecord[0] = 's' AND
     #arrRecord[1] = 'F' AND
     #arrRecord[2] = 'A') OR (#bCanActive AND
     #arrRecord[0] = 's' AND
     #arrRecord[12] = 'F' AND
     #arrRecord[13] = 'A')) THEN

     (*Get the position of the error code*)
     IF #bCanActive THEN
       #iIndex:= 15;
     ELSE
       #iIndex:= 4;
     END_IF;

     "SICK_GetValue"(iTelegramLength:= INT_TO_UINT(#fbCCom.ReqLength),
                     iValueLength:= 0,
                     nValue=> #nFncValue,
                     nErrorCode=> #nFncErrorCode,
                     iPosition:= #iIndex,
                     arrData:= #arrRecord);

     IF #nFncErrorCode = 16#0000 THEN
       #nTempErrorCode.%W1:= DWORD_TO_WORD(#nFncValue);
       #nTempErrorCode.%W0:= 16#0011; (*Error: Device error*)
     ELSE
       #nTempErrorCode.%W1:= #nFncErrorCode;
       #nTempErrorCode.%W0:= 16#0012; (*Error: SICK_GetValue error*)      
     END_IF;
   END_IF;

   (*Error detected*)
   IF #nTempErrorCode <>16#0000_0000 THEN
     RETURN;
   END_IF;


   (*================================= START REQUEST (STEP 1) =================================*)
   IF NOT #bReqBusyMem AND #bTriggerReq THEN
     #ReqDone:= false;
     #ReqBusy:= true;
     #bReqBusyMem:= true;
     #Error:= false;
     #Errorcode:= 16#0000_0000;
     #bDeviceState:= false;
     #bEnforceLogout:= false;

     (*Save the current bit selection for the job*)
     #arrSelection[0]:= #TriggerOn;
     #arrSelection[1]:= #TriggerOff;
     #arrSelection[2]:= #Matchcode;
     #arrSelection[3]:= #SavePermanent;
     #arrSelection[4]:= #ComTest;
     #arrSelection[5]:= #FreeCommand;

     (*Check CAN-ID*)
     IF #CANId > 63 THEN
       #nTempErrorCode:= 16#0000_0014; (*Error invalid CAN Id*)  
     ELSIF #CANId = 0 THEN
       #bCanActive:= false;
       #iStep:= 3; (*Check parameter input*)
     ELSE
       #bCanActive:= true;
       #iStep:= 2; (*Add CAN identifier*)
     END_IF;
   END_IF;


   (*=============================== ADD CAN IDENTIFIER (STEP 2) ==============================*)
   IF #iStep =2 THEN
     Strg_TO_Chars(Strg:= 's{ 00 01 ', pChars:= 0, Cnt=> #iIndex, Chars:=#arrCommand);

     "SICK_SetValue"(bAddBlank:= false,
                     nValue:= #CANId,
                     arrData=> #arrCommand,
                     nErrorCode=> #nFncErrorCode,
                     iPosition:= #iIndex);
     IF #nFncErrorCode <> 16#0000 THEN
       #nTempErrorCode.%W1:= #nFncErrorCode;
       #nTempErrorCode.%W0:= 16#0013; (*Error: SICK_SetValue error*)
     ELSE
       #arrCommand[#iIndex]:= '}';
       #iStep:= 3; (*Check parameter input*)
     END_IF;
   END_IF;


   (*============================= CHECK PARAMETER INPUT (STEP 3) =============================*)
   IF #iStep =3 THEN
     #iTemp1:= 0; (*Counts up the active bit selection*)

     (*Command: Trigger On*)
     IF #arrSelection[0] THEN
       #iTemp1:= #iTemp1+1;
       #iCommandIndex:= 0; (*Send a "Trigger On" command*)
     END_IF;

     (*Command: Trigger Off*)
     IF #arrSelection[1] THEN
       #iTemp1:= #iTemp1+1;
       #iCommandIndex:= 1; (*Send a "Trigger Off" command*)
     END_IF;

     (*Command: Matchcode*)
     IF #arrSelection[2] THEN
       #iTemp1:= #iTemp1+1;

       IF #Data.Matchcode.sName = '' THEN
         #nTempErrorCode:= 16#0000_0022; (*Error: Matchcode name is empty*)
       ELSIF #Data.Matchcode.nCodeType <='$20' OR #Data.Matchcode.nCodeType > '$7E' THEN
         #nTempErrorCode:= 16#0000_0023; (*Error: Invalid code type*)
       END_IF;

       #iCommandIndex:= 10; (*Send a "Login" command*)
     END_IF;

     (*Command: Save permanent*)
     IF #arrSelection[3] THEN 
       #iTemp1:= #iTemp1+1;
       #iCommandIndex:= 10; (*Send a "Login" command*)  
     END_IF;

     (*Command: Communication test*)
     IF #arrSelection[4] THEN
       #iTemp1:= #iTemp1+1;
       #iCommandIndex:= 4; (*Send a "Comm Test" command*)
     END_IF;

     (*Command: Free command*)
     IF #arrSelection[5] THEN
       #iTemp1:= #iTemp1+1;

       (*Check length*)
       IF #bCanActive THEN
         #iTemp2:= INT_TO_UDINT(LEN(#Data.FreeCommand.sCommand))+11;
       ELSE
         #iTemp2:= INT_TO_UDINT(LEN(#Data.FreeCommand.sCommand));
       END_IF;

       IF (LEN(#Data.FreeCommand.sCommand) <=0) OR (#iTemp2 > #iCommandSize) THEN
         #nTempErrorCode:= 16#0000_0020; (*Error: Invalid free command length*)
       END_IF;

       #iCommandIndex:= 5; (*Send a "Free Command" command*)
     END_IF;

     (*Check bit sum of the command selection*)
     IF #iTemp1 <>1 THEN
       #nTempErrorCode:= 16#0000_0015; (*Error: More than one or no parameter selected*)   
     END_IF;

     (*Check if a error was detected*)
     IF #nTempErrorCode = 16#0000_0000 THEN
       #iStep:= 4; (*Create CoLa command*)
     END_IF;
   END_IF;


   (*============================== CREATE COLA COMMAND (STEP 4) ==============================*)
   IF #iStep =4 THEN
     CASE #iCommandIndex OF

     (*Create "Trigger On" command*)
     0:  IF #bCanActive THEN
           Strg_TO_Chars(Strg:= 'MN mTCgateon', pChars:= 12, Cnt=> #iTemp3, Chars:=#arrCommand);
           #iCommandLength:= UDINT_TO_UINT(#iTemp3)+12;
         ELSE
           Strg_TO_Chars(Strg:= 'sMN mTCgateon', pChars:= 0, Cnt=> #iTemp3, Chars:=#arrCommand);
           #iCommandLength:= UDINT_TO_UINT(#iTemp3);
         END_IF;
         #iStep:= 5; (*Send command*)

     (*Create "Trigger Off" command*)
     1:  IF #bCanActive THEN
           Strg_TO_Chars(Strg:= 'MN mTCgateoff', pChars:= 12, Cnt=> #iTemp3, Chars:=#arrCommand);
           #iCommandLength:= UDINT_TO_UINT(#iTemp3)+12;
         ELSE
           Strg_TO_Chars(Strg:= 'sMN mTCgateoff', pChars:= 0, Cnt=> #iTemp3, Chars:=#arrCommand);
           #iCommandLength:= UDINT_TO_UINT(#iTemp3);
         END_IF;
         #iStep:= 5; (*Send command*)

     (*Create "Matchcode" command*)
     2:  IF #bCanActive THEN
           Strg_TO_Chars(Strg:= 'MN mEVSetMatchCode 00 ', pChars:= 12, Cnt=> #iTemp3, Chars:=#arrCommand);
           #iIndex:= UDINT_TO_UINT(#iTemp3+12);
         ELSE
           Strg_TO_Chars(Strg:= 'sMN mEVSetMatchCode 00 ', pChars:= 0, Cnt=> #iTemp3, Chars:=#arrCommand);
           #iIndex:= UDINT_TO_UINT(#iTemp3);
         END_IF;

         (*Add matchcode name*)
         Strg_TO_Chars(Strg:= CONCAT(IN1:= 'name="', IN2:= #Data.Matchcode.sName), pChars:= #iIndex, Cnt=> #iTemp3, Chars:=#arrCommand);
         #iIndex:= #iIndex+UDINT_TO_UINT(#iTemp3);

         (*Add codeType*)
         Strg_TO_Chars(Strg:= '" codeType="', pChars:= #iIndex, Cnt=> #iTemp3, Chars:=#arrCommand);
         #iIndex:= #iIndex+UDINT_TO_UINT(#iTemp3);
         IF #Data.Matchcode.nCodeType = '*' THEN
           Strg_TO_Chars(Strg:= 'dontCare', pChars:= #iIndex, Cnt=> #iTemp3, Chars:=#arrCommand);
           #iIndex:= #iIndex+UDINT_TO_UINT(#iTemp3);
         ELSE
           #arrCommand[#iIndex]:= #Data.Matchcode.nCodeType;
           #iIndex:= #iIndex+1;
         END_IF;

         (*Add Min/Max length*)
         Strg_TO_Chars(Strg:= '" length="', pChars:= #iIndex, Cnt=> #iTemp3, Chars:=#arrCommand);
         #iIndex:= #iIndex+UDINT_TO_UINT(#iTemp3);
         IF #Data.Matchcode.iMinMaxLength = 0 THEN
           Strg_TO_Chars(Strg:= 'dontCare', pChars:= #iIndex, Cnt=> #iTemp3, Chars:=#arrCommand);
           #iIndex:= #iIndex+UDINT_TO_UINT(#iTemp3);
         ELSE
           #arrCommand[#iIndex]:= ((#Data.Matchcode.iMinMaxLength/100) MOD 10)+16#30;     
           #arrCommand[#iIndex+1]:= ((#Data.Matchcode.iMinMaxLength/10) MOD 10)+16#30;
           #arrCommand[#iIndex+2]:= (#Data.Matchcode.iMinMaxLength MOD 10)+16#30;
           #iIndex:= #iIndex+3;
         END_IF;

         (*Add content*)
         Strg_TO_Chars(Strg:= CONCAT(IN1:= '" content="', IN2:= #Data.Matchcode.sContent), pChars:= #iIndex, Cnt=> #iTemp3, Chars:=#arrCommand);
         #iIndex:= #iIndex+UDINT_TO_UINT(#iTemp3);
         #arrCommand[#iIndex]:= '"';


         (*Overwrite the matchcode length*)
         IF #bCanActive THEN
           #nFncValue:= #iIndex-33;      (*Length of the #Matchcode command*)
           #iCommandLength:= #iIndex+1;  (*Length of the whole CoLa command*)
           #iIndex:= 31;                 (*Startindex of the matchcode length*)
         ELSE
           #nFncValue:= #iIndex-22;      (*Length of the #Matchcode command*)
           #iCommandLength:= #iIndex+1;  (*Length of the whole CoLa command*)
           #iIndex:= 20;                 (*Startindex of the matchcode length*)
         END_IF;

         "SICK_SetValue"(bAddBlank:= false,
                         nValue:= #nFncValue,
                         arrData=> #arrCommand,
                         nErrorCode=> #nFncErrorCode,
                         iPosition:=#iIndex);
         IF #nFncErrorCode <> 16#0000 THEN
           #nTempErrorCode.%W1:= #nFncErrorCode;
           #nTempErrorCode.%W0:= 16#0013; (*Error: SICK_SetValue error*)
         ELSE
           #iStep:= 5; (*Send command*)
         END_IF;

     (*Create "Save Permanent" command*)   
     3:  IF #bCanActive THEN
           Strg_TO_Chars(Strg:= 'MN mEEwriteall', pChars:= 12, Cnt=> #iTemp3, Chars:=#arrCommand);
           #iCommandLength:= UDINT_TO_UINT(#iTemp3+12);
         ELSE
           Strg_TO_Chars(Strg:= 'sMN mEEwriteall', pChars:= 0, Cnt=> #iTemp3, Chars:=#arrCommand);
           #iCommandLength:= UDINT_TO_UINT(#iTemp3);
         END_IF;
         #iStep:= 5; (*Send command*)

     (*Create "Communication Test" command*)
     4:  IF #bCanActive THEN
           Strg_TO_Chars(Strg:= 'RI0', pChars:= 12, Cnt=> #iTemp3, Chars:=#arrCommand);
           #iCommandLength:= UDINT_TO_UINT(#iTemp3)+12;
         ELSE
           Strg_TO_Chars(Strg:= 'sRI0', pChars:= 0, Cnt=> #iTemp3, Chars:=#arrCommand);
           #iCommandLength:= UDINT_TO_UINT(#iTemp3);
         END_IF;
         #iStep:= 5; (*Send command*)

     (*Create "Free Command"*)
     5:  IF #bCanActive THEN
           Strg_TO_Chars(Strg:= DELETE(IN:= #Data.FreeCommand.sCommand, L:=1, P:=1), pChars:= 12, Cnt=> #iTemp3, Chars:=#arrCommand);
           #iCommandLength:= UDINT_TO_UINT(#iTemp3)+12;
         ELSE
           Strg_TO_Chars(Strg:= #Data.FreeCommand.sCommand, pChars:= 0, Cnt=> #iTemp3, Chars:=#arrCommand);
           #iCommandLength:= UDINT_TO_UINT(#iTemp3);
         END_IF;
         #iStep:= 5; (*Send command*)

     (*Create "Login" command*)
     10: IF #bCanActive THEN
           Strg_TO_Chars(Strg:= 'MN SetAccessMode 03 F4724744', pChars:= 12, Cnt=> #iTemp3, Chars:=#arrCommand);
           #iCommandLength:= UDINT_TO_UINT(#iTemp3)+12;
         ELSE
           Strg_TO_Chars(Strg:= 'sMN SetAccessMode 03 F4724744', pChars:= 0, Cnt=> #iTemp3, Chars:=#arrCommand);
           #iCommandLength:= UDINT_TO_UINT(#iTemp3);
         END_IF;
         #iStep:= 5; (*Send command*)

     (*Create "Logout" command*)
     11: IF #bCanActive THEN
           Strg_TO_Chars(Strg:= 'MN Run', pChars:= 12, Cnt=> #iTemp3, Chars:=#arrCommand);
           #iCommandLength:= UDINT_TO_UINT(#iTemp3)+12;
         ELSE
           Strg_TO_Chars(Strg:= 'sMN Run', pChars:= 0, Cnt=> #iTemp3, Chars:=#arrCommand);
           #iCommandLength:= UDINT_TO_UINT(#iTemp3);
         END_IF;
         #iStep:= 5; (*Send command*)

       END_CASE;
   END_IF;


   (*=============================== SEND COLA COMMAND (STEP 5) ===============================*)
   IF #iStep =5 THEN
     IF NOT #fbCCom.ReqBusy AND NOT #bTriggerDone AND NOT #bTriggerError THEN
       #fbCCom.Req:= true;
       #iStep:= 6; (*Wait for the command answer*)
     END_IF;
   END_IF;


   (*========================== WAIT FOR THE COMMAND ANSWER (STEP 6) ==========================*)
   IF #iStep =6 THEN
     (*Communication error*)
     IF #bTriggerError THEN
       #nTempErrorCode:= #fbCCom.Errorcode; (*Error: Communication error*)

       (*Communication done*)
     ELSIF #bTriggerDone THEN
       #iStep:= 7; (*Check the command answer*)
     END_IF;
   END_IF;


   (*============================= CHECK COMMAND RESPONSE (STEP 7) ============================*)
   IF #iStep =7 THEN
     CASE #iCommandIndex OF

     (*Check "Trigger On" response*)
     0:  IF #bCanActive THEN
           IF #arrRecord[0] = 's' AND
             #arrRecord[12] = 'A' AND
             #arrRecord[13] = 'N' AND
             #arrRecord[22] = 'o' AND
             #arrRecord[23] = 'n' AND
             #arrRecord[24] = ' ' AND
             #arrRecord[25] = '1' THEN

             #iStep:= 8; (*Action performed*)
           ELSE
             #nTempErrorCode:= 16#0000_0016; (*Error: Invalid device answer*)                    
           END_IF;
         ELSE
           IF #arrRecord[0] = 's' AND
             #arrRecord[1] = 'A' AND
             #arrRecord[2] = 'N' AND
             #arrRecord[11] = 'o' AND
             #arrRecord[12] = 'n' AND
             #arrRecord[13] = ' ' AND
             #arrRecord[14] = '1' THEN

             #iStep:= 8; (*Action performed*)
           ELSE
             #nTempErrorCode:= 16#0000_0016; (*Error: Invalid device answer*)        
           END_IF;
         END_IF;

     (*Check "Trigger Off" response*)
     1:  IF #bCanActive THEN
           IF #arrRecord[0] = 's' AND
             #arrRecord[12] = 'A' AND
             #arrRecord[13] = 'N' AND
             #arrRecord[22] = 'o' AND
             #arrRecord[23] = 'f' AND
             #arrRecord[24] = 'f' AND
             #arrRecord[25] = ' ' AND
             #arrRecord[26] = '1' THEN

             #iStep:= 8; (*Action performed*)
           ELSE
             #nTempErrorCode:= 16#0000_0016; (*Error: Invalid device answer*)          
           END_IF;
         ELSE
           IF #arrRecord[0] = 's' AND
             #arrRecord[1] = 'A' AND
             #arrRecord[2] = 'N' AND
             #arrRecord[11] = 'o' AND
             #arrRecord[12] = 'f' AND
             #arrRecord[13] = 'f' AND
             #arrRecord[14] = ' ' AND
             #arrRecord[15] = '1' THEN

             #iStep:= 8; (*Action performed*)
           ELSE  
             #nTempErrorCode:= 16#0000_0016; (*Error: Invalid device answer*)          
           END_IF;
         END_IF;

     (*Check "Matchcode" response*)
     2:  IF #bCanActive THEN
           IF NOT(#arrRecord[0] = 's' AND
             #arrRecord[12] = 'A' AND
             #arrRecord[13] = 'N' AND
             #arrRecord[27] = 'o' AND
             #arrRecord[28] = 'd' AND
             #arrRecord[29] = 'e' AND
             #arrRecord[30] = ' ' AND
             #arrRecord[31] = '1') THEN

             #nTempErrorCode:= 16#0000_0016; (*Error: Invalid device answer*)          
           END_IF;
         ELSE
           IF NOT(#arrRecord[0] = 's' AND
             #arrRecord[1] = 'A' AND
             #arrRecord[2] = 'N' AND
             #arrRecord[16] = 'o' AND
             #arrRecord[17] = 'd' AND
             #arrRecord[18] = 'e' AND
             #arrRecord[19] = ' ' AND
             #arrRecord[20] = '1') THEN

             #nTempErrorCode:= 16#0000_0016; (*Error: Invalid device answer*)          
           END_IF;
         END_IF;

         IF #nTempErrorCode = 0 THEN
           #iCommandIndex:= 11; (*Logout*)
           #iStep:= 4;         (*Create command*)
         END_IF;    

     (*Check "Save Permanent" response*)
     3:  IF #bCanActive THEN
           IF NOT(#arrRecord[0] = 's' AND
             #arrRecord[12] = 'A' AND
             #arrRecord[13] = 'N' AND
             #arrRecord[23] = 'a' AND
             #arrRecord[24] = 'l' AND
             #arrRecord[25] = 'l' AND
             #arrRecord[26] = ' ' AND
             #arrRecord[27] = '1') THEN

             #nTempErrorCode:= 16#0000_0016; (*Error: Invalid device answer*)          
           END_IF;
         ELSE
           IF NOT(#arrRecord[0] = 's' AND
             #arrRecord[1] = 'A' AND
             #arrRecord[2] = 'N' AND
             #arrRecord[12] = 'a' AND
             #arrRecord[13] = 'l' AND
             #arrRecord[14] = 'l' AND
             #arrRecord[15] = ' ' AND
             #arrRecord[16] = '1') THEN

             #nTempErrorCode:= 16#0000_0016; (*Error: Invalid device answer*)          
           END_IF;
         END_IF;

         IF #nTempErrorCode = 0 THEN
           #iCommandIndex:= 11; (*Logout*)
           #iStep:= 4;         (*Create command*)
         END_IF;

     (*Check "Communication Test" response*)
     4:  IF #bCanActive THEN
           IF #arrRecord[0] = 's' AND
             #arrRecord[12] = 'R' AND
             #arrRecord[13] = 'A' AND
             #arrRecord[14] = ' ' THEN

             #iStep:= 8; (*Action performed*)
           ELSE
             #nTempErrorCode:= 16#0000_0016; (*Error: Invalid device answer*)          
           END_IF;
         ELSE
           IF #arrRecord[0] = 's' AND
             #arrRecord[1] = 'R' AND
             #arrRecord[2] = 'A' AND
             #arrRecord[3] = ' ' THEN

             #iStep:= 8; (*Action performed*)
           ELSE  
             #nTempErrorCode:= 16#0000_0016; (*Error: Invalid device answer*)          
           END_IF;
         END_IF;

     (*Check "Free command" response*)
     5:  IF #fbCCom.ReqLength <= MAX_LEN(#Data.FreeCommand.sResult) THEN 
           Chars_TO_Strg(Chars:= #arrRecord, pChars:= 0, Cnt:= INT_TO_UINT(#fbCCom.ReqLength),Strg=> #Data.FreeCommand.sResult);
           #iStep:= 8; (*Action performed*)
         ELSE
           #nTempErrorCode:= 16#0000_0021; (*Error: Free command result > Result string*)
         END_IF;

     (*Check "Login" response*)
     10:  IF #bCanActive THEN
           IF NOT(#arrRecord[0] = 's' AND
             #arrRecord[12] = 'A' AND
             #arrRecord[13] = 'N' AND
             #arrRecord[24] = 'M' AND
             #arrRecord[25] = 'o' AND
             #arrRecord[26] = 'd' AND
             #arrRecord[27] = 'e' AND
             #arrRecord[28] = ' ' AND
             #arrRecord[29] = '1') THEN

             #nTempErrorCode:= 16#0000_0016; (*Error: Invalid device answer*)          
           END_IF;
         ELSE
           IF NOT(#arrRecord[0] = 's' AND
             #arrRecord[1] = 'A' AND
             #arrRecord[2] = 'N' AND
             #arrRecord[13] = 'M' AND
             #arrRecord[14] = 'o' AND
             #arrRecord[15] = 'd' AND
             #arrRecord[16] = 'e' AND
             #arrRecord[17] = ' ' AND
             #arrRecord[18] = '1') THEN

             #nTempErrorCode:= 16#0000_0016; (*Error: Invalid device answer*)          
           END_IF;
         END_IF;

         IF #nTempErrorCode = 0 THEN
           IF #arrSelection[2] THEN
             #iCommandIndex:= 2; (*Matchcode*)
             #iStep:= 4;         (*Create command*)
           ELSIF #arrSelection[3] THEN
             #iCommandIndex:= 3; (*Save permanent*)
             #iStep:= 4;         (*Create command*)       
           END_IF;
           #bDeviceState:= true; (*Edit-Mode active*)
         END_IF;

     (*Check "Logout" response*)
     11:  IF #bCanActive THEN
           IF #arrRecord[0] = 's' AND
             #arrRecord[12] = 'A' AND
             #arrRecord[13] = 'N' AND
             #arrRecord[14] = ' ' AND
             #arrRecord[15] = 'R' AND
             #arrRecord[16] = 'u' AND
             #arrRecord[17] = 'n' AND
             #arrRecord[18] = ' ' AND
             #arrRecord[19] = '1' THEN

             #bDeviceState:= false; (*Run-Mode active*)
             #iStep:= 8; (*Action performed*)
           ELSE
             #nTempErrorCode:= 16#0000_0016; (*Error: Invalid device answer*)          
           END_IF;
         ELSE
           IF #arrRecord[0] = 's' AND
             #arrRecord[1] = 'A' AND
             #arrRecord[2] = 'N' AND
             #arrRecord[3] = ' ' AND
             #arrRecord[4] = 'R' AND
             #arrRecord[5] = 'u' AND
             #arrRecord[6] = 'n' AND
             #arrRecord[7] = ' ' AND
             #arrRecord[8] = '1' THEN

             #bDeviceState:= false; (*Run-Mode active*)
             #iStep:= 8; (*Action performed*)
           ELSE  
             #nTempErrorCode:= 16#0000_0016; (*Error: Invalid device answer*)          
           END_IF;
         END_IF;
     END_CASE;
   END_IF;


   (*================================ ACTION PERFORMED (STEP 8) ===============================*)
   IF #iStep =8 THEN
     IF #bEnforceLogout THEN
       #nTempErrorCode:= #nLogoutErrorCode;
     ELSE
       #ReqDone:= true;
       #ReqBusy:= false;
       #bReqBusyMem:= false;
       #iStep:= 0;
     END_IF;
   END_IF;


   (*====================================== COMMUNICATION =====================================*)
   #fbCCom(HWInputIdent:= #HWInputIdent,
           HWInputLength:= #HWInputLength,
           HWOutputIdent:= #HWOutputIdent,
           HWOutputLength:= #HWOutputLength,
           TOut:= #TOut+T#1s,
           CommandLength:= #iCommandLength,
           arrCommand:= #arrCommand,
           arrRecord:= #arrRecord);

   (*Reset the request flag every cycle*)
   #fbCCom.Req:= false;

   (*Read result error*)
   IF #fbCCom.RdLength <0 AND #fbCCom.RdDone THEN
     #Data.ReadingResult.iLength:= -1; (*Error: Reading result longer than record array*)
     FOR #iTemp1:= 1 TO UINT_TO_INT(#iReadingResultSize) DO
       #Data.ReadingResult.arrResult[#iTemp1]:= 16#00;
     END_FOR;

   (*Handling of the reading result*)
   ELSIF #fbCCom.RdDone THEN
     IF #fbCCom.RdLength > #iReadingResultSize THEN
       #Data.ReadingResult.iLength:= -1; (*Error: Reading result longer than reading result array*)
       FOR #iTemp1:= 1 TO UINT_TO_INT(#iReadingResultSize) DO
         #Data.ReadingResult.arrResult[#iTemp1]:= 16#00;
       END_FOR;
     ELSE
       MOVE_BLK(IN:= #arrRecord[0], COUNT:= INT_TO_UINT(#fbCCom.RdLength), OUT=> #Data.ReadingResult.arrResult[1]);
       IF (#Data.ReadingResult.iCounter >=255) THEN
         #Data.ReadingResult.iCounter:= 0;
       ELSE
         #Data.ReadingResult.iCounter:= #Data.ReadingResult.iCounter+1;
       END_IF;
       #Data.ReadingResult.iLength:= #fbCCom.RdLength;
       #RdDone:= true;
     END_IF;
   END_IF;
END_FUNCTION_BLOCK

FUNCTION_BLOCK "SICK_CCOMM_PNDP"   // FB10, SCL
TITLE = SICK_CCOM_PNDP
{ S7_Optimized_Access := 'TRUE' }
AUTHOR : SICKAG
FAMILY : Ident
VERSION : 1.2
// The function block use a Profinet/Probibus connection to communicate with a SICK AutoIdent
// device. The FB makes it possible to send and receive sensor data. The Confirmed Messaging 
// protocol (CM-Protocol) is used to receive even long fragmented read results.
// stored: AutoNumber false, IsIECCheckEnabled false, IsRetainMemResEnabled false, MemoryReserve 100, SetENOAutomatically false, UDAEnableTagReadback false
   VAR_INPUT
      HWInputIdent : HW_IO;   // Hardware identification number of the input module
      HWInputLength : USInt;   // Size of the input module
      HWOutputIdent : HW_IO;   // Hardware identification number of the output module
      HWOutputLength : USInt;   // Size of the output module
      TOut : Time := T#5s;   // Time out
      Req : Bool;   // A positive edge starts the request
      CommandLength : UInt;   // Byte length of the command
   END_VAR
   VAR_OUTPUT
      RdDone : Bool;   // Reading result arrived
      RdLength : Int;   // Byte length of the reading result
      ReqDone : Bool;   // Requested data available
      ReqBusy : Bool;   // Request busy
      ReqLength : Int;   // Byte length of the requested data
      Error : Bool;   // Error
      Errorcode : DWord;   // Error code
   END_VAR
   VAR_IN_OUT
      arrCommand : Array[0..499] of Byte;
      arrRecord : Array[0..499] of Byte;
   END_VAR
   VAR
      bTriggerReq { ExternalAccessible := 'False'; ExternalVisible := 'False'; ExternalWritable := 'False'} : Bool := false;   // Rising edge detection
      bTriggerReqMem { ExternalAccessible := 'False'; ExternalVisible := 'False'; ExternalWritable := 'False'} : Bool := false;   // Rising edge detection
      bReadFrag { ExternalAccessible := 'False'; ExternalVisible := 'False'; ExternalWritable := 'False'} : Bool;
      bWriteFrag { ExternalAccessible := 'False'; ExternalVisible := 'False'; ExternalWritable := 'False'} : Bool;
      bReqBusyMem : Bool;
      iReadStep { ExternalAccessible := 'False'; ExternalVisible := 'False'; ExternalWritable := 'False'} : USInt;
      iWriteStep { ExternalAccessible := 'False'; ExternalVisible := 'False'; ExternalWritable := 'False'} : USInt;
      iReadIndex { ExternalAccessible := 'False'; ExternalVisible := 'False'; ExternalWritable := 'False'} : UInt;
      iWriteIndex { ExternalAccessible := 'False'; ExternalVisible := 'False'; ExternalWritable := 'False'} : UInt;
      iReadHeaderLength { ExternalAccessible := 'False'; ExternalVisible := 'False'; ExternalWritable := 'False'} : UInt;
      iWriteHeaderLength { ExternalAccessible := 'False'; ExternalVisible := 'False'; ExternalWritable := 'False'} : UInt;
      iReadFragmentLength { ExternalAccessible := 'False'; ExternalVisible := 'False'; ExternalWritable := 'False'} : UInt;
      iWriteFragmentLength { ExternalAccessible := 'False'; ExternalVisible := 'False'; ExternalWritable := 'False'} : UInt;
      iRecordSize { ExternalAccessible := 'False'; ExternalVisible := 'False'; ExternalWritable := 'False'} : UInt;
      iCommandSize { ExternalAccessible := 'False'; ExternalVisible := 'False'; ExternalWritable := 'False'} : UInt;
      nTempErrorCode { ExternalAccessible := 'False'; ExternalVisible := 'False'; ExternalWritable := 'False'} : DWord;
      arrInputImage : Array[0..127] of Byte;
      arrOutputImage : Array[0..127] of Byte;
      fbTimeout { ExternalAccessible := 'False'; ExternalVisible := 'False'; ExternalWritable := 'False'; S7_SetPoint := 'True'} : TON_TIME;
   END_VAR
   VAR_TEMP
      iTemp1 : Int;
      iTemp2 : UDInt;
      iTemp3 : UDInt;
   END_VAR
BEGIN
   (*===========================================================================================
   Name:   SICK_CCOMM_PNDP
   Author: SICK AG
   =============================================================================================
   Description: 
   The function block use a Profinet/Probibus connection to communicate with a SICK AutoIdent
   device. The FB makes it possible to send and receive sensor data. The Confirmed Messaging 
   protocol (CM-Protocol) is used to receive even long fragmented read results.

   Send a command:
   The "Req" parameter must be triggered with a rising edge (signal change FALSE to TRUE) in 
   order to carry out the function. For the time during which a valid response has yet to be 
   received from the device, the "ReqBusy" parameter is used to signal  that a response is still 
   pending. The module signals the "ReqDone" = TRUE output parameter when the function has been 
   successfully completed. If data was requested by the device, this data is copied into the 
   Record (arrRecord). The "ReqDone" indicates that new data has been received  for a PLC cycle.
   Only one CoLa-A command request can be send to the same device at one time. 

   Receive a reading result:
   Data sent via trigger command or directly by the device (e.g., direct trigger via a light 
   barrier) is stored in the Record (arrRecord). The "RdDone" output indicates that new data 
   has been received for a PLC cycle. The data sent by the device can be changed or adapted in 
   output format of SOPAS-ET. 

   This AOI supports the folowing SICK devices:
   - Lector6xx
   - RFU6xx
   - CLV6xx 
   - RFH6xx
   =============================================================================================
   Confirmed Messaging Protocol definitions:
   arrInputImage[0]        = Status byte 
   arrInputImage[1]        = Receive counter
   arrInputImage[2]        = Transmit counter back
   arrInputImage[3]        = Command length LSB
   arrInputImage[4]        = Command length MSB
   arrInputImage[5..127]   = Device response (CoLa-A)

   arrOutputImage[0]       = Status byte 
   arrOutputImage[1]       = Receive counter back
   arrOutputImage[2]       = Transmit counter
   arrOutputImage[3]       = Command length LSB
   arrOutputImage[4]       = Command length MSB
   arrOutputImage[5..127]  = Device request (CoLa-A)
   =============================================================================================
   Version history:
   Date       | Version | Created under               | Author  | Remark
   ---------------------------------------------------------------------------------------------
   16/01/2014 | V1.0    | TIA Portal V12 SP1 Update 2 | SICK AG | Initial version
   07/08/2014 | V1.1    | TIA Portal V12 SP1 Update 4 | SICK AG | Replace R_TRIG function 
   22/04/2015 | V1.2    | TIA Portal V12 SP1 Update 4 | SICK AG | Avoid warnings that occur with 
                                                                  TIA V13
   ============================================================================================*)

   (*===================================== INITIALISATION =====================================*)
   #iRecordSize:= 500;   (*Length of the arrRecord array*)
   #iCommandSize:= 500;  (*Length of the arrCommand array*)

   #RdDone:= false;
   #iReadStep:= 0;

   (*Rising edge detection of the request flag*)
   #bTriggerReq:= #Req AND NOT #bTriggerReqMem;
   #bTriggerReqMem:= #Req;

   (*Error detection*)
   IF #nTempErrorCode <>16#0000_0000 THEN
     #ReqDone:= false;
     #ReqBusy:= false;
     #bReqBusyMem:= false;
     #Error:= true;
     #Errorcode:= #nTempErrorCode;
     #nTempErrorCode:= 16#0000_0000;
     #ReqLength:= 0;
     #iWriteStep:= 0;
     RETURN;
   END_IF;

   (*Time out detection*)
   #fbTimeout(IN:=#bReqBusyMem, PT:=#TOut);
   IF #fbTimeout.Q THEN
     #nTempErrorCode:= 16#0000_0001; (*Error: Time out*) 
   END_IF;

   (*Check the hardware ident length of the input module*)
   IF #HWInputLength <8 OR #HWInputLength >128 THEN
     #nTempErrorCode:= 16#0000_0002; (*Error: Incorrect module input length*)
   END_IF;

   (*Check the hardware ident length of the output module*)
   IF #HWOutputLength <8 OR #HWOutputLength >128 THEN
     #nTempErrorCode:= 16#0000_0003; (*Error: Incorrect module output length*)
   END_IF;

   (*Error detected*)
   IF #nTempErrorCode <>16#0000_0000 THEN
     RETURN;
   END_IF;


   (*===================================== COMMUNICATION ======================================*)
   (*Set output data*)
   #iTemp1:= DPWR_DAT(LADDR:= #HWOutputIdent, RECORD:= #arrOutputImage);
   IF #iTemp1 <>0 THEN
     #nTempErrorCode.%W1:= #iTemp1;
     #nTempErrorCode.%W0:= 16#0004; (*Error: Set output data via DPWR_DAT*)
     RETURN;
   END_IF;

   (*Get input data*)
   #iTemp1:= DPRD_DAT(LADDR:= #HWInputIdent, RECORD=> #arrInputImage);
   IF #iTemp1 <>0 THEN
     #nTempErrorCode.%W1:= #iTemp1;
     #nTempErrorCode.%W0:= 16#0005; (*Error: Get input data via DPRD_DAT*)
     RETURN;
   END_IF;

   (*Receive counter ==0 && Receive counter back <>0*)
   IF #arrInputImage[1] =0 AND #arrOutputImage[1] <>0 THEN
     #arrOutputImage[1]:= #arrInputImage[1]; (*Recive counter => Receive counter back*)
     RETURN;
   END_IF;

   (*Transmit counter <> Transmit counter back*)
   IF NOT #bReqBusyMem AND (#arrInputImage[2] <> #arrOutputImage[2]) THEN
     #arrOutputImage[2]:= 0; (*0 => Transmit counter*)
     RETURN;
   END_IF;


   (*============================== HANDLING OF THE RECEIVED DATA =============================*)
   (*New telegram available*)
   IF NOT (#arrInputImage[1] = #arrOutputImage[1]) THEN

     (*Reset error every incoming telegram (Read only mode, e.g. for hand held scanners)*)
     IF #CommandLength <=0 THEN
       #Error:= false;
       #Errorcode:= 16#0000_0000;
     END_IF;

     (*Confirm the receive counter*)
     #arrOutputImage[1]:= #arrInputImage[1];

     (*Get telegram length from the received header*)
     #iReadHeaderLength.%B0:= #arrInputImage[3];
     #iReadHeaderLength.%B1:= #arrInputImage[4];

     (*Check if fragmentation is not active at the moment*)
     IF NOT #bReadFrag THEN
       #iReadIndex:= 0;

       (*Check if fragmentation is needed*)
       IF (#HWInputLength-5) < #iReadHeaderLength THEN
         #bReadFrag:= true;
       END_IF;
     END_IF;

     (*Fragmentation is needed*)
     IF #bReadFrag THEN
       IF (#HWInputLength-5) < #iReadHeaderLength THEN
         #iReadFragmentLength:= #HWInputLength-5;
       ELSE
         #iReadFragmentLength:= #iReadHeaderLength;
       END_IF;

     (*No fragmentation needed*)
     ELSE
       #iReadFragmentLength:= #iReadHeaderLength;
     END_IF;

     (*Copy input data into the output record*)
     IF (#iReadIndex+#iReadFragmentLength) <= #iRecordSize THEN
       MOVE_BLK(IN:= #arrInputImage[5], COUNT:= #iReadFragmentLength, OUT=> #arrRecord[#iReadIndex]);
     END_IF;

     (*Check if all data has been received*)
     IF (#HWInputLength-5) < #iReadHeaderLength THEN
       #iReadIndex:= #iReadIndex+#iReadFragmentLength;

     (*All data has been received*)
     ELSE
       #bReadFrag:= false;
       #iReadStep:= 1;
     END_IF;

     (*Incoming data filter*)
     (* - Check if the receiving telegram os a CoLa answer on a requested 
          comand or a reading result.

         sRA  sWA  sMA  sAN  sAI  sEA  sPX  s{   sSI  sSN  sFA
     sRN  X                                       X    X    X
     sRI  X                                       X    X    X
     sWN       X                                  X    X    X
     sWI       X                                  X    X    X
     sMN            X    X                        X    X    X
     sMI            X         X                   X    X    X
     sEN                           X              X    X    X
     sEI                           X              X    X    X
     sPE                                X         X    X    X
     s{                                      X    X    X    X
     *)
     IF #iReadStep =1 THEN
       (*Filter is only active, while requested data expected*)
       IF #bReqBusyMem THEN
         IF #CommandLength >3 THEN
           (*Get the prefix from the requested command (e.g. 'sRN '*)   
           #iTemp2.%B3:= #arrCommand[0];
           #iTemp2.%B2:= #arrCommand[1];
           #iTemp2.%B1:= #arrCommand[2];
           #iTemp2.%B0:= 16#20;

           (*Get the prefix from the command response (e.g. 'sRA ')*)
           #iTemp3.%B3:= #arrRecord[0];
           #iTemp3.%B2:= #arrRecord[1];
           #iTemp3.%B1:= #arrRecord[2];
           #iTemp3.%B0:= 16#20;
         ELSE
           #iTemp2:= 16#0000_0000;
           #iTemp3:= 16#0000_0000;
         END_IF;

         CASE #iTemp3 OF
         (*'s{  '*)
         16#737B2020:  IF #iTemp2 = 16#737B2020 THEN
                         #iReadStep:= 2; (*Command response*)
                       ELSE
                         #iReadStep:= 3; (*Reading result*)
                       END_IF;

         (*'sRA '*)
         16#73524120:  IF (#iTemp2 = 16#73524E20) OR (#iTemp2 = 16#73524920) THEN
                         #iReadStep:= 2; (*Command response*)
                       ELSE
                         #iReadStep:= 3; (*Reading result*)
                       END_IF;

         (*'sWA '*)
         16#73574120:  IF (#iTemp2 = 16#73574E20) OR (#iTemp2 = 16#73574920) THEN
                         #iReadStep:= 2; (*Command response*)
                       ELSE
                         #iReadStep:= 3; (*Reading result*)
                       END_IF;

         (*'sMA '*)
         16#734D4120:  IF (#iTemp2 = 16#734D4E20) OR (#iTemp2 = 16#734D4920) THEN
                         #iReadStep:= 2; (*Command response*)
                       ELSE
                         #iReadStep:= 3; (*Reading result*)
                       END_IF;

         (*'sAN '*)
         16#73414E20:  IF #iTemp2 = 16#734D4E20 THEN
                         #iReadStep:= 2; (*Command response*)
                       ELSE
                         #iReadStep:= 3; (*Reading result*)
                       END_IF;

         (*'sAI '*)
         16#73414920:  IF #iTemp2 = 16#734D4920 THEN
                         #iReadStep:= 2; (*Command response*)
                       ELSE
                         #iReadStep:= 3; (*Reading result*)
                       END_IF;

         (*'sEA '*)
         16#73454120:  IF (#iTemp2 = 16#73454E20) OR (#iTemp2 = 16#73454920) THEN
                         #iReadStep:= 2; (*Command response*)
                       ELSE
                         #iReadStep:= 3; (*Reading result*)
                       END_IF;

         (*'sPX '*)
         16#73505820:  IF #iTemp2 = 16#73504520 THEN
                         #iReadStep:= 2; (*Command response*)
                       ELSE
                         #iReadStep:= 3; (*Reading result*)
                       END_IF;

         (*'sSI '*)
         16#73534920:  #iReadStep:= 3; (*Reading result*)

         (*'sSN '*)
         16#73534E20:  #iReadStep:= 3; (*Reading result*)

         (*'sFA '*)
         16#73464120:  #iReadStep:= 2; (*Command response*)

         (*Invalid CoLa-A answer*)
         ELSE
           (*Check if a user defined command is used (Request == Response)*)
           FOR #iTemp1:= 0 TO UINT_TO_INT(#CommandLength-1) DO
             IF #arrCommand[#iTemp1] = #arrRecord[#iTemp1] THEN
               #iReadStep:= 2; (*Command response*)
             ELSE
               #iReadStep:= 3; (*Reading result*)
               EXIT;
             END_IF;
           END_FOR;
         END_CASE;

       (*Reading result*)
       ELSE
         #iReadStep:= 3;  (*Reading result*)
       END_IF;
     END_IF;

     (*Incoming telegram is a command response*)
     IF #iReadStep =2 THEN
       IF (#iReadIndex+#iReadFragmentLength) <= #iRecordSize THEN
         #ReqLength:= UDINT_TO_INT(#iReadIndex+#iReadFragmentLength);
         #ReqDone:= true;
         #ReqBusy:= false;
         #bReqBusyMem:= false;
       ELSE
         #nTempErrorCode:= 16#0000_0006; (*Error: Incoming command response > Record size*)
       END_IF;
     END_IF;

     (*Incoming telegram is a reading result*)
     IF #iReadStep =3 THEN
       IF (#iReadIndex+#iReadFragmentLength) <= #iRecordSize THEN
         #RdLength:= UDINT_TO_INT(#iReadIndex+#iReadFragmentLength);
         #RdDone:= true;
       ELSE
         #RdLength:= -1;
         #RdDone:= false;    
       END_IF;
     END_IF;
   END_IF;


   (*=========================== HANDLING OF THE DATA TO BE WRITTEN ===========================*)
   IF #bTriggerReq AND NOT #bReqBusyMem THEN
     #ReqDone:= false;
     #ReqBusy:= true;
     #bReqBusyMem:= true;
     #Error:= false;
     #Errorcode:= 16#0000_0000;
     #iWriteIndex:= 0;

     (*Check command length*)
     IF #CommandLength <=0 THEN
       #nTempErrorCode:= 16#0000_0007; (*Error: Command length <= 0*)
       RETURN;
     ELSIF #CommandLength > #iCommandSize THEN
       #nTempErrorCode:= 16#0000_0008; (*Error: Command length > command array*)
       RETURN;
     END_IF;

     (*Check if the the command telegram must be fragmented*)
     IF (#HWOutputLength-5) < #CommandLength THEN
       #iWriteFragmentLength:= #HWOutputLength-5;
     ELSE
       #iWriteFragmentLength:= #CommandLength;
     END_IF;

     #iWriteHeaderLength:= #CommandLength;
     #iWriteStep:= 1;  
   END_IF;

   (*Write step 1: Command transfer*)
   IF (#iWriteStep =1) AND(#arrInputImage[2] = #arrOutputImage[2]) THEN

     (*Copy command data into the output record*)
     IF((#iWriteIndex+#iWriteFragmentLength) <= #iCommandSize) AND (#iWriteFragmentLength <= (#HWOutputLength-5)) THEN
       MOVE_BLK(IN:= #arrCommand[#iWriteIndex], COUNT:= #iWriteFragmentLength, OUT=> #arrOutputImage[5]);
       (*Increment transmit counter*)
       IF #arrOutputImage[2] = 16#FF THEN
         #arrOutputImage[2]:= 16#01; (*Counter overflow, zero is skipped*)
       ELSE
         #arrOutputImage[2]:= #arrOutputImage[2]+1;
       END_IF;

       (*Set command/fragment length*)
       #arrOutputImage[3]:= #iWriteHeaderLength.%B0;
       #arrOutputImage[4]:= #iWriteHeaderLength.%B1;

       (*Next step*)
       #iWriteStep:= 2;
     ELSE
       #nTempErrorCode:= 16#0000_0009; (*Error: Fragmentation error*)
     END_IF;
       RETURN;
   END_IF;

   (*Write step 2: Fragmentation handling*)
   IF #iWriteStep =2 THEN

     (*Fragmentation is needed*)
     IF (#HWOutputLength-5) < #iWriteHeaderLength THEN
       #bWriteFrag:= true;

       (*Next index*)
       #iWriteIndex:= #iWriteIndex+#iWriteFragmentLength;

       (*Set next header length*)
       #iWriteHeaderLength:= #iWriteHeaderLength-#iWriteFragmentLength;

       (*Set next fragment length*)
       IF (#HWOutputLength-5) < #iWriteHeaderLength THEN
         #iWriteFragmentLength:= #HWOutputLength-5;
       ELSE
         #iWriteFragmentLength:= #iWriteHeaderLength;
       END_IF;

     (*Fragmentation is not needed*)
     ELSE
       #bWriteFrag:= false;
     END_IF;

     (*Next step*)
     #iWriteStep:= 3;
   END_IF;

   (*Write step 3: Check if the transmission of the command/fragment is done*)
   IF #iWriteStep =3 THEN

     (*Transmit counter back == Transmit counter*)
     IF #arrInputImage[2] = #arrOutputImage[2] THEN
       IF #bWriteFrag THEN
         #iWriteStep:= 1;
       ELSE
         #iWriteStep:= 0;
       END_IF;
     END_IF;
   END_IF;
END_FUNCTION_BLOCK

FUNCTION_BLOCK "SICK_Barcode_FB"   // FB19, SCL
{ S7_Optimized_Access := 'TRUE' }
VERSION : 0.1
// stored: AutoNumber true, IsIECCheckEnabled false, IsRetainMemResEnabled false, MemoryReserve 100, SetENOAutomatically false, UDAEnableTagReadback false
   VAR_INPUT
      Rd_Done : Bool;
      Req_Done : Bool;
      Req_Busy : Bool;
      Error : Bool;
      arrResult : Array[1..200] of Byte;
      iCounter : USInt;
      iLength : Int;
      Error_Code : DWord;
   END_VAR
   VAR_OUTPUT
      Test_Comm : Bool;
      Enable_Trigger : Bool;
      Disable_Trigger : Bool;
      Enable_Req : Bool;
      Result : String;
      Test_OK : Bool;
   END_VAR
BEGIN
   //Communication Test
   IF "VTD_BCD_Start_Comm_Test_HMI_Tag" THEN
       #Test_Comm := 1;
       #Enable_Req := 1;
       "IEC_Timer_0_DB_1".TON(IN:=True,
                              PT:=t#1s);
   END_IF;

   //TEST OK
   IF #Req_Done AND "IEC_Timer_0_DB_1".Q AND NOT #Error THEN
       #Test_OK := 1;
       #Test_Comm := 0;
       #Enable_Req := 0;
       "VTD_BCD_Start_Comm_Test_HMI_Tag" := 0;
       "IEC_Timer_0_DB_1".TON(IN := FALSE,
                              PT := t#0s);
   END_IF;

   //ERROR
   IF "IEC_Timer_0_DB_1".Q AND #Error THEN
           #Test_OK := 0;
           #Test_Comm := 0;
           #Enable_Req := 0;
           "VTD_BCD_Start_Comm_Test_HMI_Tag" := 0;
           "IEC_Timer_0_DB_1".TON(IN := FALSE,
                                  PT := t#0s);
       END_IF;

   //Enable Trigger
       IF "VTD_BCD_Enable_Trigger_HMI_Tag" OR "Auto_Start_Barcode" THEN
       #Enable_Trigger := 1;
       #Enable_Req := 1;
       "VTD_BCD_Disable_Trigger_HMI_Tag" := 0;
       #Disable_Trigger := 0;
   //Disable Trigger
   ELSIF "VTD_BCD_Disable_Trigger_HMI_Tag" OR "Auto_Stop_Barcode" THEN
       #Disable_Trigger := 1;
       #Enable_Req := 1;
       "VTD_BCD_Enable_Trigger_HMI_Tag" := 0;
       #Enable_Trigger := 0;
   ELSE
       #Enable_Trigger := 0;
       #Enable_Req := 0;
       #Disable_Trigger := 0;
   END_IF;


   "R_TRIG_DB_5"(CLK:=#Rd_Done);

   IF "R_TRIG_DB_5".Q OR "IEC_Timer_0_DB_18".Q OR
       ("VTD_BCD_Enable_Trigger_HMI_Tag" AND "VTD_BCD_Disable_Trigger_HMI_Tag")
   THEN
       "VTD_BCD_Disable_Trigger_HMI_Tag" := 0;
       #Enable_Trigger := 0;
       #Disable_Trigger := 0;
       #Enable_Req := 0;
       "IEC_Timer_0_DB_18".TON(IN := FALSE,
                               PT := T#0S);
       "Auto_Stop_Barcode" := 0;
   END_IF;

   "IEC_Timer_0_DB_18".TON(IN:=("VTD_BCD_Enable_Trigger_HMI_Tag" OR "VTD_BCD_Disable_Trigger_HMI_Tag" OR "Auto_Start_Barcode" OR "Auto_Stop_Barcode"),
                               PT:=T#10S);

   #Result := "ByteArrayToString_1"(Lenght := #iLength, ByteArray := #arrResult);
END_FUNCTION_BLOCK

FUNCTION "Weighing Station FC" : Void   // FC31, SCL
{ S7_Optimized_Access := 'TRUE' }
VERSION : 0.1
// stored: AutoNumber true, IsIECCheckEnabled false, SetENOAutomatically false, UDAEnableTagReadback false
   VAR_INPUT
      Start : Bool;
      MinWeight : Real;
      MaxWeight : Real;
   END_VAR
BEGIN
   "R_TRIG_DB_25"(CLK:=#Start, Q=> "R_Start_WS");

   CASE "State_WS" OF
       0: // IDLE / READY
           "Control_DB"."Weighing Station".Ready := TRUE;
           "Control_DB"."Weighing Station".Running := FALSE;
           IF "R_Start_WS" THEN
               "Control_DB"."Weighing Station".Done := FALSE;
               "Control_DB"."Weighing Station".Valid := FALSE;
               "Control_DB"."Weighing Station".Ready := FALSE;
               "Control_DB"."Weighing Station".Error_ID := 0;
               "State_WS" := 10;
           END_IF;

       10:
           "Control_DB"."Weighing Station".Start := FALSE;
           "Control_DB"."Weighing Station".Running := TRUE;
           IF "Control_DB".PopUp_Cnv[1].Inputs."Lift Up" THEN

               IF NOT "SAI_Cyclic_WeightProc_DB".DataOK THEN
                   "Control_DB"."Weighing Station".Error_ID.%X0 := TRUE;
                   "Control_DB"."Weighing Station".Done := TRUE;
                   "State_WS" := 100;
               ELSE
                   "Control_DB"."Weighing Station".Weight := "SAI_Cyclic_WeightProc_DB".RealTimeWeight;
                   "State_WS" := 20;
               END_IF;
           END_IF;
           "IEC_Timer_0_DB_17".TON(IN:=TRUE,
                                   PT:=t#10S);
           IF "IEC_Timer_0_DB_17".Q THEN
               "IEC_Timer_0_DB_17".TON(IN := FALSE,
                                       PT := t#0S);
               // "Control_DB"."Weighing Station".Done := TRUE;
               "State_WS" := 20;
           END_IF;

       20:
           IF "Control_DB"."Weighing Station".Weight < #MinWeight THEN
               "Control_DB"."Weighing Station".Valid := FALSE;
               // "Control_DB"."Weighing Station".Error_ID.%X1 := TRUE;
           ELSIF "Control_DB"."Weighing Station".Weight > #MaxWeight THEN
               "Control_DB"."Weighing Station".Valid := FALSE;
               // "Control_DB"."Weighing Station".Error_ID.%X2 := TRUE;
           ELSE
               "Control_DB"."Weighing Station".Valid := TRUE;
               "Control_DB"."Weighing Station".Error_ID := 0;
           END_IF;
           "State_WS" := 100;

       100:
           "Control_DB"."Weighing Station".Running := FALSE;
           "Control_DB"."Weighing Station".Done := TRUE;
           "State_WS" := 0;

   END_CASE;

   IF "Reset_All" THEN
       "Control_DB"."Weighing Station".Error_ID := 0;
   END_IF;
END_FUNCTION

FUNCTION "MT_ACT_Application" : Void   // FC30, LAD
{ S7_Optimized_Access := 'FALSE' }
VERSION : 0.1
// stored: AutoNumber true, IsIECCheckEnabled false, SetENOAutomatically false, UDAEnableTagReadback false
BEGIN

REGION Network 1: Cyclic Weighing Data
   // All the cyclical read and write commands can be issued from this Function Block.
   // The cyclic commands are triggered following a positive trigger. These commands are Tare Immediate, Tare Stable, Zero Immediate, Zero Stable, Pretare and Clear Tare. 
   // Upon successful execution of these commands, the DONE output bit will be set ON.
   // ERROR output bit will be set on if there is an error with the command execution.
   // Note: Only one cyclic command is possible at any one time.
   // If Net weight is required after executed a zero or tare command, insert decimal value "3" into the "WeightCmd" variable before triggering the cyclic scale command. Else, with decimal value "1" in the "WeightCmd" variable, the Function Block will return Gross Weight after the cyclic scale command. 
   // "DataOK" bit is set ON when the scale is in operation mode, not overloaded and not underload.
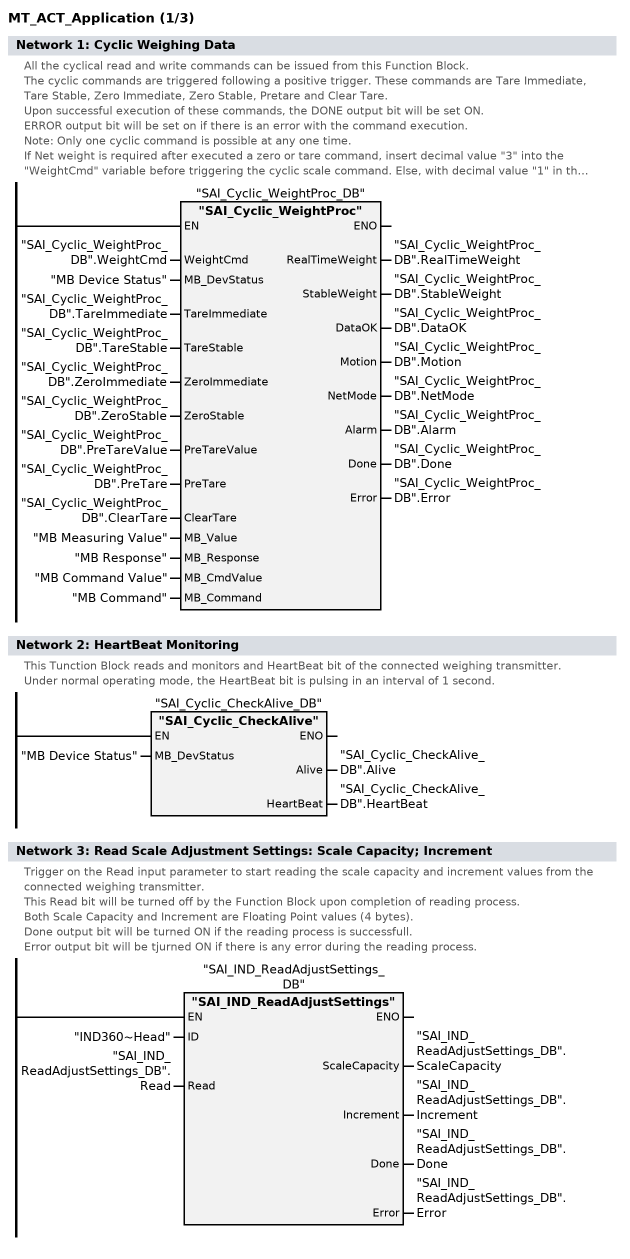
   RUNG wire#powerrail
      "SAI_Cyclic_WeightProc_DB"(WeightCmd := "SAI_Cyclic_WeightProc_DB".WeightCmd, MB_DevStatus := "MB Device Status", TareImmediate := "SAI_Cyclic_WeightProc_DB".TareImmediate, TareStable := "SAI_Cyclic_WeightProc_DB".TareStable, ZeroImmediate := "SAI_Cyclic_WeightProc_DB".ZeroImmediate, ZeroStable := "SAI_Cyclic_WeightProc_DB".ZeroStable, PreTareValue := "SAI_Cyclic_WeightProc_DB".PreTareValue, PreTare := "SAI_Cyclic_WeightProc_DB".PreTare, ClearTare := "SAI_Cyclic_WeightProc_DB".ClearTare, MB_Value := "MB Measuring Value", MB_Response := "MB Response", MB_CmdValue := "MB Command Value", MB_Command := "MB Command", RealTimeWeight => "SAI_Cyclic_WeightProc_DB".RealTimeWeight, StableWeight => "SAI_Cyclic_WeightProc_DB".StableWeight, DataOK => "SAI_Cyclic_WeightProc_DB".DataOK, Motion => "SAI_Cyclic_WeightProc_DB".Motion, NetMode => "SAI_Cyclic_WeightProc_DB".NetMode, Alarm => "SAI_Cyclic_WeightProc_DB".Alarm, Done => "SAI_Cyclic_WeightProc_DB".Done, Error => "SAI_Cyclic_WeightProc_DB".Error)
   END_RUNG
   // the same network as SCL:
   "SAI_Cyclic_WeightProc_DB"(WeightCmd := "SAI_Cyclic_WeightProc_DB".WeightCmd,   // "SAI_Cyclic_WeightProc"
                           MB_DevStatus := "MB Device Status",
                           TareImmediate := "SAI_Cyclic_WeightProc_DB".TareImmediate,
                           TareStable := "SAI_Cyclic_WeightProc_DB".TareStable,
                           ZeroImmediate := "SAI_Cyclic_WeightProc_DB".ZeroImmediate,
                           ZeroStable := "SAI_Cyclic_WeightProc_DB".ZeroStable,
                           PreTareValue := "SAI_Cyclic_WeightProc_DB".PreTareValue,
                           PreTare := "SAI_Cyclic_WeightProc_DB".PreTare,
                           ClearTare := "SAI_Cyclic_WeightProc_DB".ClearTare,
                           MB_Value := "MB Measuring Value",
                           MB_Response := "MB Response",
                           MB_CmdValue := "MB Command Value",
                           MB_Command := "MB Command",
                           RealTimeWeight => "SAI_Cyclic_WeightProc_DB".RealTimeWeight,
                           StableWeight => "SAI_Cyclic_WeightProc_DB".StableWeight,
                           DataOK => "SAI_Cyclic_WeightProc_DB".DataOK,
                           Motion => "SAI_Cyclic_WeightProc_DB".Motion,
                           NetMode => "SAI_Cyclic_WeightProc_DB".NetMode,
                           Alarm => "SAI_Cyclic_WeightProc_DB".Alarm,
                           Done => "SAI_Cyclic_WeightProc_DB".Done,
                           Error => "SAI_Cyclic_WeightProc_DB".Error);
END_REGION

REGION Network 2: HeartBeat Monitoring
   // This Tunction Block reads and monitors and HeartBeat bit of the connected weighing transmitter.
   // Under normal operating mode, the HeartBeat bit is pulsing in an interval of 1 second.
   RUNG wire#powerrail
      "SAI_Cyclic_CheckAlive_DB"(MB_DevStatus := "MB Device Status", Alive => "SAI_Cyclic_CheckAlive_DB".Alive, HeartBeat => "SAI_Cyclic_CheckAlive_DB".HeartBeat)
   END_RUNG
   // the same network as SCL:
   "SAI_Cyclic_CheckAlive_DB"(MB_DevStatus := "MB Device Status",   // "SAI_Cyclic_CheckAlive"
                           Alive => "SAI_Cyclic_CheckAlive_DB".Alive,
                           HeartBeat => "SAI_Cyclic_CheckAlive_DB".HeartBeat);
END_REGION

REGION Network 3: Read Scale Adjustment Settings: Scale Capacity; Increment
   // Trigger on the Read input parameter to start reading the scale capacity and increment values from the connected weighing transmitter.
   // This Read bit will be turned off by the Function Block upon completion of reading process.
   // Both Scale Capacity and Increment are Floating Point values (4 bytes).
   // Done output bit will be turned ON if the reading process is successfull.
   // Error output bit will be tjurned ON if there is any error during the reading process.
   RUNG wire#powerrail
      "SAI_IND_ReadAdjustSettings_DB"(ID := "IND360~Head", Read := "SAI_IND_ReadAdjustSettings_DB".Read, ScaleCapacity => "SAI_IND_ReadAdjustSettings_DB".ScaleCapacity, Increment => "SAI_IND_ReadAdjustSettings_DB".Increment, Done => "SAI_IND_ReadAdjustSettings_DB".Done, Error => "SAI_IND_ReadAdjustSettings_DB".Error)
   END_RUNG
   // the same network as SCL:
   "SAI_IND_ReadAdjustSettings_DB"(ID := "IND360~Head",   // "SAI_IND_ReadAdjustSettings"
                           Read := "SAI_IND_ReadAdjustSettings_DB".Read,
                           ScaleCapacity => "SAI_IND_ReadAdjustSettings_DB".ScaleCapacity,
                           Increment => "SAI_IND_ReadAdjustSettings_DB".Increment,
                           Done => "SAI_IND_ReadAdjustSettings_DB".Done,
                           Error => "SAI_IND_ReadAdjustSettings_DB".Error);
END_REGION

REGION Network 4: Write new Scale Adjustment Settings: Scale Capacity; Increment
   // Trigger on the Write input parameter to start writing the new scale capacity and increment settings to the connected weighing transmitter.
   // Both Scale Capacity and Increment are Floating Point values (4 bytes).
   // Make sure both settings are valid and correct before triggering the Write input bit.
   // This Write bit will be turned off by the Function Block upon completion of writing process.
   // Done output bit will be set ON if the reading process is successfull.
   // Error output bit will be set ON if there is any error during the reading process.
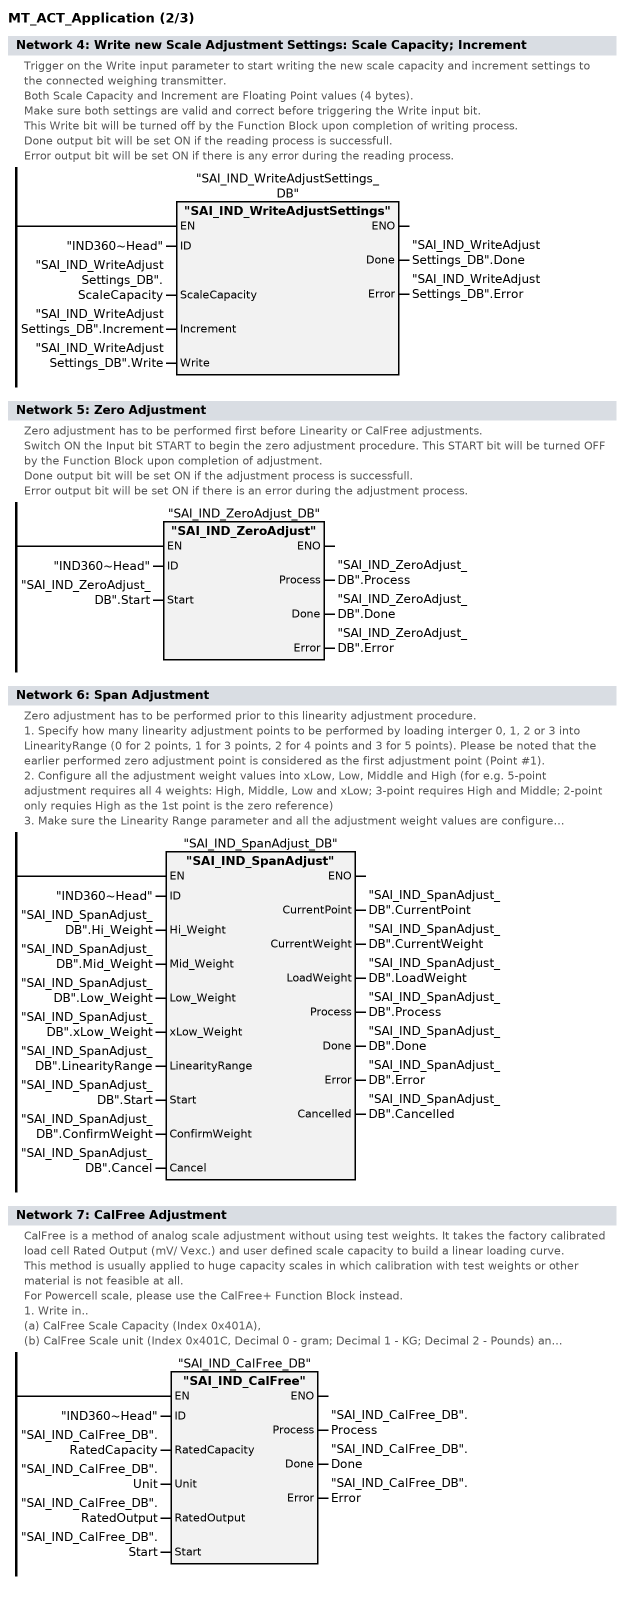
   RUNG wire#powerrail
      "SAI_IND_WriteAdjustSettings_DB"(ID := "IND360~Head", ScaleCapacity := "SAI_IND_WriteAdjustSettings_DB".ScaleCapacity, Increment := "SAI_IND_WriteAdjustSettings_DB".Increment, Write := "SAI_IND_WriteAdjustSettings_DB".Write, Done => "SAI_IND_WriteAdjustSettings_DB".Done, Error => "SAI_IND_WriteAdjustSettings_DB".Error)
   END_RUNG
   // the same network as SCL:
   "SAI_IND_WriteAdjustSettings_DB"(ID := "IND360~Head",   // "SAI_IND_WriteAdjustSettings"
                           ScaleCapacity := "SAI_IND_WriteAdjustSettings_DB".ScaleCapacity,
                           Increment := "SAI_IND_WriteAdjustSettings_DB".Increment,
                           Write := "SAI_IND_WriteAdjustSettings_DB".Write,
                           Done => "SAI_IND_WriteAdjustSettings_DB".Done,
                           Error => "SAI_IND_WriteAdjustSettings_DB".Error);
END_REGION

REGION Network 5: Zero Adjustment
   // Zero adjustment has to be performed first before Linearity or CalFree adjustments.
   // Switch ON the Input bit START to begin the zero adjustment procedure. This START bit will be turned OFF by the Function Block upon completion of adjustment. 
   // Done output bit will be set ON if the adjustment process is successfull.
   // Error output bit will be set ON if there is an error during the adjustment process.
   RUNG wire#powerrail
      "SAI_IND_ZeroAdjust_DB"(ID := "IND360~Head", Start := "SAI_IND_ZeroAdjust_DB".Start, Process => "SAI_IND_ZeroAdjust_DB".Process, Done => "SAI_IND_ZeroAdjust_DB".Done, Error => "SAI_IND_ZeroAdjust_DB".Error)
   END_RUNG
   // the same network as SCL:
   "SAI_IND_ZeroAdjust_DB"(ID := "IND360~Head",   // "SAI_IND_ZeroAdjust"
                           Start := "SAI_IND_ZeroAdjust_DB".Start,
                           Process => "SAI_IND_ZeroAdjust_DB".Process,
                           Done => "SAI_IND_ZeroAdjust_DB".Done,
                           Error => "SAI_IND_ZeroAdjust_DB".Error);
END_REGION

